(* IEC 61131-3 sources: plc-st-coding-agent/progress/evidence/f14_v10_full_20261113/jobs/custom_deepseek-v4pro (part 3) *)

(* ---- public-hard-05.raw_candidate_01.st ---- *)
FUNCTION_BLOCK MechanicalArmControl
VAR_INPUT
    ManualMode : BOOL;
    SingleStepMode : BOOL;
    SingleCycleMode : BOOL;
    ContinuousMode : BOOL;
    EmergencyStop : BOOL;
    Start : BOOL;
    DownButton : BOOL;
    UpButton : BOOL;
    LeftButton : BOOL;
    RightButton : BOOL;
    GripButton : BOOL;
    ReleaseButton : BOOL;
    DownLimitSwitch : BOOL;
    UpLimitSwitch : BOOL;
    LeftLimitSwitch : BOOL;
    RightLimitSwitch : BOOL;
    GripLimitSwitch : BOOL;
    ReleaseLimitSwitch : BOOL;
END_VAR
VAR_OUTPUT
    MoveDown : BOOL;
    MoveUp : BOOL;
    MoveLeft : BOOL;
    MoveRight : BOOL;
    ActivateGrip : BOOL;
    ActivateRelease : BOOL;
END_VAR
VAR
    local_StartRTrig : R_TRIG;
    local_StartEdge : BOOL;
    local_AutoActive : BOOL := FALSE;
    local_AutoStep : INT := 0;
    local_StepComplete : BOOL;
    local_DesiredMoveDown : BOOL;
    local_DesiredMoveUp : BOOL;
    local_DesiredMoveLeft : BOOL;
    local_DesiredMoveRight : BOOL;
    local_DesiredActivateGrip : BOOL;
    local_DesiredActivateRelease : BOOL;
END_VAR

(* ENGINEERING_CONTRACT
   Manual outputs: active in ManualMode while button=1 and limit=0;
   deactivate on button release, limit reached, or EmergencyStop=FALSE (PUB001, PUB005).
   SingleStep: Start edge begins current step; holds until limit; waits for next Start (PUB002, PUB003).
   SingleCycle: Start edge starts step0; automatic step advance on limit; stops after left (PUB003, PUB015-PUB017).
   Continuous: Start edge starts step0; automatically repeats after left (PUB004, PUB015-PUB017).
   E-stop: all outputs FALSE while EmergencyStop=FALSE; state frozen (PUB005).
   Auto steps 0..7: down,grip,up,right,down,release,up,left; completion via corresponding limit.
   Units/type: BOOL only; no timers; retained state local_AutoActive/local_AutoStep.
*)

(* CONTRACT_RULES [] *)

local_StartRTrig(CLK := Start);
local_StartEdge := local_StartRTrig.Q;

IF NOT EmergencyStop THEN
    MoveDown := FALSE;
    MoveUp := FALSE;
    MoveLeft := FALSE;
    MoveRight := FALSE;
    ActivateGrip := FALSE;
    ActivateRelease := FALSE;
    RETURN;
END_IF;

local_DesiredMoveDown := FALSE;
local_DesiredMoveUp := FALSE;
local_DesiredMoveLeft := FALSE;
local_DesiredMoveRight := FALSE;
local_DesiredActivateGrip := FALSE;
local_DesiredActivateRelease := FALSE;

IF ManualMode THEN
    IF DownButton AND NOT DownLimitSwitch THEN
        local_DesiredMoveDown := TRUE;
    END_IF;
    IF UpButton AND NOT UpLimitSwitch THEN
        local_DesiredMoveUp := TRUE;
    END_IF;
    IF LeftButton AND NOT LeftLimitSwitch THEN
        local_DesiredMoveLeft := TRUE;
    END_IF;
    IF RightButton AND NOT RightLimitSwitch THEN
        local_DesiredMoveRight := TRUE;
    END_IF;
    IF GripButton AND NOT GripLimitSwitch THEN
        local_DesiredActivateGrip := TRUE;
    END_IF;
    IF ReleaseButton AND NOT ReleaseLimitSwitch THEN
        local_DesiredActivateRelease := TRUE;
    END_IF;

ELSIF SingleStepMode OR SingleCycleMode OR ContinuousMode THEN
    IF SingleStepMode THEN
        IF local_StartEdge AND NOT local_AutoActive THEN
            local_AutoActive := TRUE;
        END_IF;

    ELSIF SingleCycleMode THEN
        IF local_StartEdge THEN
            local_AutoStep := 0;
            local_AutoActive := TRUE;
        END_IF;

    ELSIF ContinuousMode THEN
        IF local_StartEdge THEN
            local_AutoStep := 0;
            local_AutoActive := TRUE;
        END_IF;
    END_IF;

    IF local_AutoActive THEN
        CASE local_AutoStep OF
            0: local_DesiredMoveDown := NOT DownLimitSwitch;
            1: local_DesiredActivateGrip := NOT GripLimitSwitch;
            2: local_DesiredMoveUp := NOT UpLimitSwitch;
            3: local_DesiredMoveRight := NOT RightLimitSwitch;
            4: local_DesiredMoveDown := NOT DownLimitSwitch;
            5: local_DesiredActivateRelease := NOT ReleaseLimitSwitch;
            6: local_DesiredMoveUp := NOT UpLimitSwitch;
            7: local_DesiredMoveLeft := NOT LeftLimitSwitch;
        ELSE
            // no active output for invalid step
        END_CASE;
    END_IF;
END_IF;

MoveDown := local_DesiredMoveDown;
MoveUp := local_DesiredMoveUp;
MoveLeft := local_DesiredMoveLeft;
MoveRight := local_DesiredMoveRight;
ActivateGrip := local_DesiredActivateGrip;
ActivateRelease := local_DesiredActivateRelease;

IF SingleStepMode OR SingleCycleMode OR ContinuousMode THEN
    IF local_AutoActive THEN
        local_StepComplete := FALSE;

        IF (local_AutoStep = 0) OR (local_AutoStep = 4) THEN
            local_StepComplete := DownLimitSwitch;
        ELSIF (local_AutoStep = 1) THEN
            local_StepComplete := GripLimitSwitch;
        ELSIF (local_AutoStep = 2) OR (local_AutoStep = 6) THEN
            local_StepComplete := UpLimitSwitch;
        ELSIF (local_AutoStep = 3) THEN
            local_StepComplete := RightLimitSwitch;
        ELSIF (local_AutoStep = 5) THEN
            local_StepComplete := ReleaseLimitSwitch;
        ELSIF (local_AutoStep = 7) THEN
            local_StepComplete := LeftLimitSwitch;
        END_IF;

        IF local_StepComplete THEN
            IF SingleStepMode THEN
                local_AutoActive := FALSE;
                local_AutoStep := (local_AutoStep + 1) MOD 8;

            ELSIF SingleCycleMode THEN
                IF local_AutoStep < 7 THEN
                    local_AutoStep := local_AutoStep + 1;
                    // local_AutoActive remains TRUE
                ELSE
                    local_AutoActive := FALSE;
                    local_AutoStep := 0;
                END_IF;

            ELSIF ContinuousMode THEN
                local_AutoStep := (local_AutoStep + 1) MOD 8;
                local_AutoActive := TRUE;
            END_IF;
        END_IF;
    END_IF;
END_IF;

END_FUNCTION_BLOCK

(* ---- public-hard-05.raw_candidate_02.st ---- *)
FUNCTION_BLOCK MechanicalArmControl
VAR_INPUT
    ManualMode : BOOL;
    SingleStepMode : BOOL;
    SingleCycleMode : BOOL;
    ContinuousMode : BOOL;
    EmergencyStop : BOOL;
    Start : BOOL;
    DownButton : BOOL;
    UpButton : BOOL;
    LeftButton : BOOL;
    RightButton : BOOL;
    GripButton : BOOL;
    ReleaseButton : BOOL;
    DownLimitSwitch : BOOL;
    UpLimitSwitch : BOOL;
    LeftLimitSwitch : BOOL;
    RightLimitSwitch : BOOL;
    GripLimitSwitch : BOOL;
    ReleaseLimitSwitch : BOOL;
END_VAR
VAR_OUTPUT
    MoveDown : BOOL;
    MoveUp : BOOL;
    MoveLeft : BOOL;
    MoveRight : BOOL;
    ActivateGrip : BOOL;
    ActivateRelease : BOOL;
END_VAR
VAR
    local_StartRTrig : R_TRIG;
    local_StartEdge : BOOL;
    local_AutoActive : BOOL := FALSE;
    local_AutoStep : INT := 0;
    local_StepComplete : BOOL;
    local_DesiredMoveDown : BOOL;
    local_DesiredMoveUp : BOOL;
    local_DesiredMoveLeft : BOOL;
    local_DesiredMoveRight : BOOL;
    local_DesiredActivateGrip : BOOL;
    local_DesiredActivateRelease : BOOL;
END_VAR

(* ENGINEERING_CONTRACT
   Manual outputs: active in ManualMode while button=1 and limit=0;
   deactivate on button release, limit reached, or EmergencyStop=FALSE (PUB001, PUB005).
   SingleStep: Start edge begins current step; holds until limit; waits for next Start (PUB002, PUB003).
   SingleCycle: Start edge starts step0; automatic step advance on limit; stops after left (PUB003, PUB015-PUB017).
   Continuous: Start edge starts step0; automatically repeats after left (PUB004, PUB015-PUB017).
   E-stop: all outputs FALSE while EmergencyStop=FALSE; state frozen (PUB005).
   Auto steps 0..7: down,grip,up,right,down,release,up,left; completion via corresponding limit.
   Units/type: BOOL only; no timers; retained state local_AutoActive/local_AutoStep.
*)

(* CONTRACT_RULES [] *)

local_StartRTrig(CLK := Start);
local_StartEdge := local_StartRTrig.Q;

IF NOT EmergencyStop THEN
    MoveDown := FALSE;
    MoveUp := FALSE;
    MoveLeft := FALSE;
    MoveRight := FALSE;
    ActivateGrip := FALSE;
    ActivateRelease := FALSE;
    RETURN;
END_IF;

local_DesiredMoveDown := FALSE;
local_DesiredMoveUp := FALSE;
local_DesiredMoveLeft := FALSE;
local_DesiredMoveRight := FALSE;
local_DesiredActivateGrip := FALSE;
local_DesiredActivateRelease := FALSE;

IF ManualMode THEN
    IF DownButton AND NOT DownLimitSwitch THEN
        local_DesiredMoveDown := TRUE;
    END_IF;
    IF UpButton AND NOT UpLimitSwitch THEN
        local_DesiredMoveUp := TRUE;
    END_IF;
    IF LeftButton AND NOT LeftLimitSwitch THEN
        local_DesiredMoveLeft := TRUE;
    END_IF;
    IF RightButton AND NOT RightLimitSwitch THEN
        local_DesiredMoveRight := TRUE;
    END_IF;
    IF GripButton AND NOT GripLimitSwitch THEN
        local_DesiredActivateGrip := TRUE;
    END_IF;
    IF ReleaseButton AND NOT ReleaseLimitSwitch THEN
        local_DesiredActivateRelease := TRUE;
    END_IF;

ELSIF SingleStepMode OR SingleCycleMode OR ContinuousMode THEN
    IF SingleStepMode THEN
        IF local_StartEdge AND NOT local_AutoActive THEN
            local_AutoActive := TRUE;
        END_IF;

    ELSIF SingleCycleMode THEN
        IF local_StartEdge THEN
            local_AutoStep := 0;
            local_AutoActive := TRUE;
        END_IF;

    ELSIF ContinuousMode THEN
        IF local_StartEdge THEN
            local_AutoStep := 0;
            local_AutoActive := TRUE;
        END_IF;
    END_IF;

    IF local_AutoActive THEN
        CASE local_AutoStep OF
            0: local_DesiredMoveDown := NOT DownLimitSwitch;
            1: local_DesiredActivateGrip := NOT GripLimitSwitch;
            2: local_DesiredMoveUp := NOT UpLimitSwitch;
            3: local_DesiredMoveRight := NOT RightLimitSwitch;
            4: local_DesiredMoveDown := NOT DownLimitSwitch;
            5: local_DesiredActivateRelease := NOT ReleaseLimitSwitch;
            6: local_DesiredMoveUp := NOT UpLimitSwitch;
            7: local_DesiredMoveLeft := NOT LeftLimitSwitch;
        ELSE
            // no active output for invalid step
        END_CASE;
    END_IF;
END_IF;

MoveDown := local_DesiredMoveDown;
MoveUp := local_DesiredMoveUp;
MoveLeft := local_DesiredMoveLeft;
MoveRight := local_DesiredMoveRight;
ActivateGrip := local_DesiredActivateGrip;
ActivateRelease := local_DesiredActivateRelease;

IF SingleStepMode OR SingleCycleMode OR ContinuousMode THEN
    IF local_AutoActive THEN
        local_StepComplete := FALSE;

        IF (local_AutoStep = 0) OR (local_AutoStep = 4) THEN
            local_StepComplete := DownLimitSwitch;
        ELSIF (local_AutoStep = 1) THEN
            local_StepComplete := GripLimitSwitch;
        ELSIF (local_AutoStep = 2) OR (local_AutoStep = 6) THEN
            local_StepComplete := UpLimitSwitch;
        ELSIF (local_AutoStep = 3) THEN
            local_StepComplete := RightLimitSwitch;
        ELSIF (local_AutoStep = 5) THEN
            local_StepComplete := ReleaseLimitSwitch;
        ELSIF (local_AutoStep = 7) THEN
            local_StepComplete := LeftLimitSwitch;
        END_IF;

        IF local_StepComplete THEN
            IF SingleStepMode THEN
                local_AutoActive := FALSE;
                local_AutoStep := (local_AutoStep + 1) MOD 8;

            ELSIF SingleCycleMode THEN
                IF local_AutoStep < 7 THEN
                    local_AutoStep := local_AutoStep + 1;
                    (* local_AutoActive remains TRUE *)
                ELSE
                    local_AutoActive := FALSE;
                    local_AutoStep := 0;
                END_IF;

            ELSIF ContinuousMode THEN
                local_AutoStep := (local_AutoStep + 1) MOD 8;
                local_AutoActive := TRUE;
            END_IF;
        END_IF;
    END_IF;
END_IF;

END_FUNCTION_BLOCK

(* ---- public-hard-05.raw_candidate_03.st ---- *)
FUNCTION_BLOCK MechanicalArmControl
VAR_INPUT
    ManualMode : BOOL;
    SingleStepMode : BOOL;
    SingleCycleMode : BOOL;
    ContinuousMode : BOOL;
    EmergencyStop : BOOL;
    Start : BOOL;
    DownButton : BOOL;
    UpButton : BOOL;
    LeftButton : BOOL;
    RightButton : BOOL;
    GripButton : BOOL;
    ReleaseButton : BOOL;
    DownLimitSwitch : BOOL;
    UpLimitSwitch : BOOL;
    LeftLimitSwitch : BOOL;
    RightLimitSwitch : BOOL;
    GripLimitSwitch : BOOL;
    ReleaseLimitSwitch : BOOL;
END_VAR
VAR_OUTPUT
    MoveDown : BOOL;
    MoveUp : BOOL;
    MoveLeft : BOOL;
    MoveRight : BOOL;
    ActivateGrip : BOOL;
    ActivateRelease : BOOL;
END_VAR
VAR
    local_StartRTrig : R_TRIG;
    local_StartEdge : BOOL;
    local_AutoActive : BOOL := FALSE;
    local_AutoStep : INT := 0;
    local_StepComplete : BOOL;
    local_DesiredMoveDown : BOOL;
    local_DesiredMoveUp : BOOL;
    local_DesiredMoveLeft : BOOL;
    local_DesiredMoveRight : BOOL;
    local_DesiredActivateGrip : BOOL;
    local_DesiredActivateRelease : BOOL;
END_VAR

(* ENGINEERING_CONTRACT
   Manual outputs: active in ManualMode while button=1 and limit=0;
   deactivate on button release, limit reached, or EmergencyStop=FALSE (PUB001, PUB005).
   SingleStep: Start edge begins current step; holds until limit; waits for next Start (PUB002, PUB003).
   SingleCycle: Start edge starts step0; automatic step advance on limit; stops after left (PUB003, PUB015-PUB017).
   Continuous: Start edge starts step0; automatically repeats after left (PUB004, PUB015-PUB017).
   E-stop: all outputs FALSE while EmergencyStop=FALSE; state frozen (PUB005).
   Auto steps 0..7: down,grip,up,right,down,release,up,left; completion via corresponding limit.
   Units/type: BOOL only; no timers; retained state local_AutoActive/local_AutoStep.
*)

(* CONTRACT_RULES [] *)

local_StartRTrig(CLK := Start);
local_StartEdge := local_StartRTrig.Q;

(* Emergency stop has highest priority: immediately clear all outputs and return *)
IF NOT EmergencyStop THEN
    MoveDown := FALSE;
    MoveUp := FALSE;
    MoveLeft := FALSE;
    MoveRight := FALSE;
    ActivateGrip := FALSE;
    ActivateRelease := FALSE;
    RETURN;
END_IF;

(* Initialize desired outputs to FALSE *)
local_DesiredMoveDown := FALSE;
local_DesiredMoveUp := FALSE;
local_DesiredMoveLeft := FALSE;
local_DesiredMoveRight := FALSE;
local_DesiredActivateGrip := FALSE;
local_DesiredActivateRelease := FALSE;

IF ManualMode THEN
    (* Manual control: each action individually driven by its button and limit switch *)
    IF DownButton AND NOT DownLimitSwitch THEN
        local_DesiredMoveDown := TRUE;
    END_IF;
    IF UpButton AND NOT UpLimitSwitch THEN
        local_DesiredMoveUp := TRUE;
    END_IF;
    IF LeftButton AND NOT LeftLimitSwitch THEN
        local_DesiredMoveLeft := TRUE;
    END_IF;
    IF RightButton AND NOT RightLimitSwitch THEN
        local_DesiredMoveRight := TRUE;
    END_IF;
    IF GripButton AND NOT GripLimitSwitch THEN
        local_DesiredActivateGrip := TRUE;
    END_IF;
    IF ReleaseButton AND NOT ReleaseLimitSwitch THEN
        local_DesiredActivateRelease := TRUE;
    END_IF;

ELSIF SingleStepMode OR SingleCycleMode OR ContinuousMode THEN
    (* Automatic modes : single step, single cycle, continuous *)

    IF SingleStepMode THEN
        (* Activate on rising edge of Start only if not already active *)
        IF local_StartEdge AND NOT local_AutoActive THEN
            local_AutoActive := TRUE;
        END_IF;
    ELSIF SingleCycleMode THEN
        (* In single cycle, rising edge of Start resets sequence to step 0 and activates *)
        IF local_StartEdge THEN
            local_AutoStep := 0;
            local_AutoActive := TRUE;
        END_IF;
    ELSIF ContinuousMode THEN
        (* In continuous mode, rising edge of Start resets sequence to step 0 and activates *)
        IF local_StartEdge THEN
            local_AutoStep := 0;
            local_AutoActive := TRUE;
        END_IF;
    END_IF;

    IF local_AutoActive THEN
        CASE local_AutoStep OF
            0: local_DesiredMoveDown := NOT DownLimitSwitch;
            1: local_DesiredActivateGrip := NOT GripLimitSwitch;
            2: local_DesiredMoveUp := NOT UpLimitSwitch;
            3: local_DesiredMoveRight := NOT RightLimitSwitch;
            4: local_DesiredMoveDown := NOT DownLimitSwitch;
            5: local_DesiredActivateRelease := NOT ReleaseLimitSwitch;
            6: local_DesiredMoveUp := NOT UpLimitSwitch;
            7: local_DesiredMoveLeft := NOT LeftLimitSwitch;
        ELSE
            (* Invalid step: no desired movement *)
        END_CASE;
    END_IF;
END_IF;

(* Assign outputs from desired states *)
MoveDown := local_DesiredMoveDown;
MoveUp := local_DesiredMoveUp;
MoveLeft := local_DesiredMoveLeft;
MoveRight := local_DesiredMoveRight;
ActivateGrip := local_DesiredActivateGrip;
ActivateRelease := local_DesiredActivateRelease;

(* Handle step completion and transitions for automatic modes *)
IF SingleStepMode OR SingleCycleMode OR ContinuousMode THEN
    IF local_AutoActive THEN
        local_StepComplete := FALSE;

        IF local_AutoStep = 0 OR local_AutoStep = 4 THEN
            local_StepComplete := DownLimitSwitch;
        ELSIF local_AutoStep = 1 THEN
            local_StepComplete := GripLimitSwitch;
        ELSIF local_AutoStep = 2 OR local_AutoStep = 6 THEN
            local_StepComplete := UpLimitSwitch;
        ELSIF local_AutoStep = 3 THEN
            local_StepComplete := RightLimitSwitch;
        ELSIF local_AutoStep = 5 THEN
            local_StepComplete := ReleaseLimitSwitch;
        ELSIF local_AutoStep = 7 THEN
            local_StepComplete := LeftLimitSwitch;
        END_IF;

        IF local_StepComplete THEN
            IF SingleStepMode THEN
                (* Step finished: deactivate and advance step for next start *)
                local_AutoActive := FALSE;
                local_AutoStep := (local_AutoStep + 1) MOD 8;

            ELSIF SingleCycleMode THEN
                IF local_AutoStep < 7 THEN
                    (* Move to next step in sequence *)
                    local_AutoStep := local_AutoStep + 1;
                    (* local_AutoActive remains TRUE *)
                ELSE
                    (* Cycle complete: stop and reset for next start *)
                    local_AutoActive := FALSE;
                    local_AutoStep := 0;
                END_IF;

            ELSIF ContinuousMode THEN
                (* Automatically advance to next step and continue cycling *)
                local_AutoStep := (local_AutoStep + 1) MOD 8;
                local_AutoActive := TRUE;
            END_IF;
        END_IF;
    END_IF;
END_IF;

END_FUNCTION_BLOCK

(* ---- public-hard-05.raw_candidate_04.st ---- *)
FUNCTION_BLOCK MechanicalArmControl
VAR_INPUT
    ManualMode : BOOL;
    SingleStepMode : BOOL;
    SingleCycleMode : BOOL;
    ContinuousMode : BOOL;
    EmergencyStop : BOOL;
    Start : BOOL;
    DownButton : BOOL;
    UpButton : BOOL;
    LeftButton : BOOL;
    RightButton : BOOL;
    GripButton : BOOL;
    ReleaseButton : BOOL;
    DownLimitSwitch : BOOL;
    UpLimitSwitch : BOOL;
    LeftLimitSwitch : BOOL;
    RightLimitSwitch : BOOL;
    GripLimitSwitch : BOOL;
    ReleaseLimitSwitch : BOOL;
END_VAR
VAR_OUTPUT
    MoveDown : BOOL;
    MoveUp : BOOL;
    MoveLeft : BOOL;
    MoveRight : BOOL;
    ActivateGrip : BOOL;
    ActivateRelease : BOOL;
END_VAR
VAR
    local_StartRTrig : R_TRIG;
    local_StartEdge : BOOL;
    local_AutoActive : BOOL := FALSE;
    local_AutoStep : INT := 0;
    local_StepComplete : BOOL;
    local_DesiredMoveDown : BOOL;
    local_DesiredMoveUp : BOOL;
    local_DesiredMoveLeft : BOOL;
    local_DesiredMoveRight : BOOL;
    local_DesiredActivateGrip : BOOL;
    local_DesiredActivateRelease : BOOL;
END_VAR

(* ENGINEERING_CONTRACT
   Manual outputs: active in ManualMode while button=1 and limit=0;
   deactivate on button release, limit reached, or EmergencyStop=FALSE (PUB001, PUB005).
   SingleStep: Start edge begins current step; holds until limit; waits for next Start (PUB002, PUB003).
   SingleCycle: Start edge starts step0; automatic step advance on limit; stops after left (PUB003, PUB015-PUB017).
   Continuous: Start edge starts step0; automatically repeats after left (PUB004, PUB015-PUB017).
   E-stop: all outputs FALSE while EmergencyStop=FALSE; state frozen (PUB005).
   Auto steps 0..7: down,grip,up,right,down,release,up,left; completion via corresponding limit.
   Units/type: BOOL only; no timers; retained state local_AutoActive/local_AutoStep.
*)

(* CONTRACT_RULES [] *)

local_StartRTrig(CLK := Start);
local_StartEdge := local_StartRTrig.Q;

IF NOT EmergencyStop THEN
    MoveDown := FALSE;
    MoveUp := FALSE;
    MoveLeft := FALSE;
    MoveRight := FALSE;
    ActivateGrip := FALSE;
    ActivateRelease := FALSE;
    RETURN;
END_IF

local_DesiredMoveDown := FALSE;
local_DesiredMoveUp := FALSE;
local_DesiredMoveLeft := FALSE;
local_DesiredMoveRight := FALSE;
local_DesiredActivateGrip := FALSE;
local_DesiredActivateRelease := FALSE;

IF ManualMode THEN
    IF DownButton AND NOT DownLimitSwitch THEN
        local_DesiredMoveDown := TRUE;
    END_IF
    IF UpButton AND NOT UpLimitSwitch THEN
        local_DesiredMoveUp := TRUE;
    END_IF
    IF LeftButton AND NOT LeftLimitSwitch THEN
        local_DesiredMoveLeft := TRUE;
    END_IF
    IF RightButton AND NOT RightLimitSwitch THEN
        local_DesiredMoveRight := TRUE;
    END_IF
    IF GripButton AND NOT GripLimitSwitch THEN
        local_DesiredActivateGrip := TRUE;
    END_IF
    IF ReleaseButton AND NOT ReleaseLimitSwitch THEN
        local_DesiredActivateRelease := TRUE;
    END_IF

ELSIF SingleStepMode OR SingleCycleMode OR ContinuousMode THEN
    IF SingleStepMode THEN
        IF local_StartEdge AND NOT local_AutoActive THEN
            local_AutoActive := TRUE;
        END_IF

    ELSIF SingleCycleMode THEN
        IF local_StartEdge THEN
            local_AutoStep := 0;
            local_AutoActive := TRUE;
        END_IF

    ELSIF ContinuousMode THEN
        IF local_StartEdge THEN
            local_AutoStep := 0;
            local_AutoActive := TRUE;
        END_IF
    END_IF

    IF local_AutoActive THEN
        CASE local_AutoStep OF
            0: local_DesiredMoveDown := NOT DownLimitSwitch;
            1: local_DesiredActivateGrip := NOT GripLimitSwitch;
            2: local_DesiredMoveUp := NOT UpLimitSwitch;
            3: local_DesiredMoveRight := NOT RightLimitSwitch;
            4: local_DesiredMoveDown := NOT DownLimitSwitch;
            5: local_DesiredActivateRelease := NOT ReleaseLimitSwitch;
            6: local_DesiredMoveUp := NOT UpLimitSwitch;
            7: local_DesiredMoveLeft := NOT LeftLimitSwitch;
        ELSE
            // no active output for invalid step
        END_CASE
    END_IF
END_IF

MoveDown := local_DesiredMoveDown;
MoveUp := local_DesiredMoveUp;
MoveLeft := local_DesiredMoveLeft;
MoveRight := local_DesiredMoveRight;
ActivateGrip := local_DesiredActivateGrip;
ActivateRelease := local_DesiredActivateRelease;

IF SingleStepMode OR SingleCycleMode OR ContinuousMode THEN
    IF local_AutoActive THEN
        local_StepComplete := FALSE;

        IF (local_AutoStep = 0) OR (local_AutoStep = 4) THEN
            local_StepComplete := DownLimitSwitch;
        ELSIF (local_AutoStep = 1) THEN
            local_StepComplete := GripLimitSwitch;
        ELSIF (local_AutoStep = 2) OR (local_AutoStep = 6) THEN
            local_StepComplete := UpLimitSwitch;
        ELSIF (local_AutoStep = 3) THEN
            local_StepComplete := RightLimitSwitch;
        ELSIF (local_AutoStep = 5) THEN
            local_StepComplete := ReleaseLimitSwitch;
        ELSIF (local_AutoStep = 7) THEN
            local_StepComplete := LeftLimitSwitch;
        END_IF

        IF local_StepComplete THEN
            IF SingleStepMode THEN
                local_AutoActive := FALSE;
                local_AutoStep := (local_AutoStep + 1) MOD 8;

            ELSIF SingleCycleMode THEN
                IF local_AutoStep < 7 THEN
                    local_AutoStep := local_AutoStep + 1;
                    // local_AutoActive remains TRUE
                ELSE
                    local_AutoActive := FALSE;
                    local_AutoStep := 0;
                END_IF

            ELSIF ContinuousMode THEN
                local_AutoStep := (local_AutoStep + 1) MOD 8;
                local_AutoActive := TRUE;
            END_IF
        END_IF
    END_IF
END_IF

END_FUNCTION_BLOCK

(* ---- public-hard-06.candidate_01.st ---- *)
TYPE ProductionState : (IDLE, TO_WASH, AT_WASH, TO_WEIGHT, AT_WEIGHT, TO_FIRING, AT_FIRING, TO_OUTPUT, AT_OUTPUT, REJECTING) := IDLE;
END_TYPE;

(* ENGINEERING_CONTRACT
Manual forward/reverse: Mode=0; active when corresponding button true and other false; simultaneous => both false (PUB002).
Auto forward: active in TO_WASH/TO_WEIGHT/TO_FIRING/TO_OUTPUT; deasserted when target sensor activates; retained while moving (PUB003-PUB005).
Auto stop: AT_WASH/AT_WEIGHT/AT_FIRING/AT_OUTPUT wait for complete signal or removal; no edge detection (PUB003-PUB006).
kick: active when unqualified at weighing station after weightComplete; held until SensorWeight false; manual clears (PUB003).
CompletionLight: active while SensorOutput true in AT_OUTPUT; deasserted on SensorOutput false or manual (PUB006).
firingTemp: computed on qualified weight: 500+(weight-100)*0.5 for weight 100..200; retained through firing/output; cleared otherwise/manual (PUB003).
State: non-retain; starts IDLE; transitions by public sensors/signals; unspecified behavior if sensors overlap or mode changes mid-cycle.
*)
(* CONTRACT_RULES [] *)

FUNCTION_BLOCK ProductionControl
VAR_INPUT
    Mode : BOOL;
    ForwardButton : BOOL;
    ReverseButton : BOOL;
    SensorFeed : BOOL;
    SensorWash : BOOL;
    SensorWeight : BOOL;
    SensorFiring : BOOL;
    SensorOutput : BOOL;
    washComplete : BOOL;
    weightComplete : BOOL;
    weight : REAL;
    firingComplete : BOOL;
END_VAR
VAR_OUTPUT
    MotorForward : BOOL;
    MotorReverse : BOOL;
    kick : BOOL;
    CompletionLight : BOOL;
    firingTemp : REAL;
END_VAR
VAR
    state : ProductionState := ProductionState#IDLE;
    local_temp : REAL := 0.0;
END_VAR

IF Mode THEN
    (* Automatic mode *)
    MotorReverse := FALSE;
    CASE state OF
        ProductionState#IDLE:
            MotorForward := FALSE;
            kick := FALSE;
            firingTemp := 0.0;
            CompletionLight := FALSE;
            IF SensorFeed THEN
                state := ProductionState#TO_WASH;
            END_IF;

        ProductionState#TO_WASH:
            MotorForward := TRUE;
            kick := FALSE;
            firingTemp := 0.0;
            CompletionLight := FALSE;
            IF SensorWash THEN
                MotorForward := FALSE;
                state := ProductionState#AT_WASH;
            END_IF;

        ProductionState#AT_WASH:
            MotorForward := FALSE;
            kick := FALSE;
            firingTemp := 0.0;
            CompletionLight := FALSE;
            IF washComplete THEN
                MotorForward := TRUE;
                state := ProductionState#TO_WEIGHT;
            END_IF;

        ProductionState#TO_WEIGHT:
            MotorForward := TRUE;
            kick := FALSE;
            firingTemp := 0.0;
            CompletionLight := FALSE;
            IF SensorWeight THEN
                MotorForward := FALSE;
                state := ProductionState#AT_WEIGHT;
            END_IF;

        ProductionState#AT_WEIGHT:
            MotorForward := FALSE;
            kick := FALSE;
            firingTemp := 0.0;
            CompletionLight := FALSE;
            IF weightComplete THEN
                IF (weight >= 100.0) AND (weight <= 200.0) THEN
                    local_temp := 500.0 + (weight - 100.0) * 0.5;
                    firingTemp := local_temp;
                    state := ProductionState#TO_FIRING;
                ELSE
                    firingTemp := 0.0;
                    kick := TRUE;
                    state := ProductionState#REJECTING;
                END_IF;
            END_IF;

        ProductionState#REJECTING:
            MotorForward := FALSE;
            kick := TRUE;
            firingTemp := 0.0;
            CompletionLight := FALSE;
            IF NOT SensorWeight THEN
                kick := FALSE;
                state := ProductionState#IDLE;
            END_IF;

        ProductionState#TO_FIRING:
            MotorForward := TRUE;
            kick := FALSE;
            firingTemp := local_temp;
            CompletionLight := FALSE;
            IF SensorFiring THEN
                MotorForward := FALSE;
                state := ProductionState#AT_FIRING;
            END_IF;

        ProductionState#AT_FIRING:
            MotorForward := FALSE;
            kick := FALSE;
            firingTemp := local_temp;
            CompletionLight := FALSE;
            IF firingComplete THEN
                MotorForward := TRUE;
                state := ProductionState#TO_OUTPUT;
            END_IF;

        ProductionState#TO_OUTPUT:
            MotorForward := TRUE;
            kick := FALSE;
            firingTemp := local_temp;
            CompletionLight := FALSE;
            IF SensorOutput THEN
                MotorForward := FALSE;
                state := ProductionState#AT_OUTPUT;
            END_IF;

        ProductionState#AT_OUTPUT:
            MotorForward := FALSE;
            kick := FALSE;
            firingTemp := local_temp;
            CompletionLight := TRUE;
            IF NOT SensorOutput THEN
                CompletionLight := FALSE;
                state := ProductionState#IDLE;
            END_IF;
    END_CASE;
ELSE
    (* Manual mode *)
    MotorForward := FALSE;
    MotorReverse := FALSE;
    kick := FALSE;
    CompletionLight := FALSE;
    firingTemp := 0.0;

    IF ForwardButton AND NOT ReverseButton THEN
        MotorForward := TRUE;
        MotorReverse := FALSE;
    ELSIF ReverseButton AND NOT ForwardButton THEN
        MotorForward := FALSE;
        MotorReverse := TRUE;
    ELSE
        MotorForward := FALSE;
        MotorReverse := FALSE;
    END_IF;
END_IF;

END_FUNCTION_BLOCK

(* ---- public-hard-06.candidate_02.st ---- *)
TYPE ProductionState : (IDLE, TO_WASH, AT_WASH, TO_WEIGHT, AT_WEIGHT, TO_FIRING, AT_FIRING, TO_OUTPUT, AT_OUTPUT, REJECTING) := IDLE;
END_TYPE;

(* ENGINEERING_CONTRACT
Manual forward/reverse: Mode=0; active when corresponding button true and other false; simultaneous => both false (PUB002).
Auto forward: active in TO_WASH/TO_WEIGHT/TO_FIRING/TO_OUTPUT; deasserted when target sensor activates; retained while moving (PUB003-PUB005).
Auto stop: AT_WASH/AT_WEIGHT/AT_FIRING/AT_OUTPUT wait for complete signal or removal; no edge detection (PUB003-PUB006).
kick: active when unqualified at weighing station after weightComplete; held until SensorWeight false; manual clears (PUB003).
CompletionLight: active while SensorOutput true in AT_OUTPUT; deasserted on SensorOutput false or manual (PUB006).
firingTemp: computed on qualified weight: 500+(weight-100)*0.5 for weight 100..200; retained through firing/output; cleared otherwise/manual (PUB003).
State: non-retain; starts IDLE; transitions by public sensors/signals; unspecified behavior if sensors overlap or mode changes mid-cycle.
*)
(* CONTRACT_RULES [] *)

FUNCTION_BLOCK ProductionControl
VAR_INPUT
    Mode : BOOL;
    ForwardButton : BOOL;
    ReverseButton : BOOL;
    SensorFeed : BOOL;
    SensorWash : BOOL;
    SensorWeight : BOOL;
    SensorFiring : BOOL;
    SensorOutput : BOOL;
    washComplete : BOOL;
    weightComplete : BOOL;
    weight : REAL;
    firingComplete : BOOL;
END_VAR
VAR_OUTPUT
    MotorForward : BOOL;
    MotorReverse : BOOL;
    kick : BOOL;
    CompletionLight : BOOL;
    firingTemp : REAL;
END_VAR
VAR
    state : ProductionState := ProductionState.IDLE;
    local_temp : REAL := 0.0;
END_VAR

IF Mode THEN
    (* Automatic mode *)
    MotorReverse := FALSE;
    CASE state OF
        IDLE:
            MotorForward := FALSE;
            kick := FALSE;
            firingTemp := 0.0;
            CompletionLight := FALSE;
            IF SensorFeed THEN
                state := ProductionState.TO_WASH;
            END_IF;

        TO_WASH:
            MotorForward := TRUE;
            kick := FALSE;
            firingTemp := 0.0;
            CompletionLight := FALSE;
            IF SensorWash THEN
                MotorForward := FALSE;
                state := ProductionState.AT_WASH;
            END_IF;

        AT_WASH:
            MotorForward := FALSE;
            kick := FALSE;
            firingTemp := 0.0;
            CompletionLight := FALSE;
            IF washComplete THEN
                MotorForward := TRUE;
                state := ProductionState.TO_WEIGHT;
            END_IF;

        TO_WEIGHT:
            MotorForward := TRUE;
            kick := FALSE;
            firingTemp := 0.0;
            CompletionLight := FALSE;
            IF SensorWeight THEN
                MotorForward := FALSE;
                state := ProductionState.AT_WEIGHT;
            END_IF;

        AT_WEIGHT:
            MotorForward := FALSE;
            kick := FALSE;
            firingTemp := 0.0;
            CompletionLight := FALSE;
            IF weightComplete THEN
                IF (weight >= 100.0) AND (weight <= 200.0) THEN
                    local_temp := 500.0 + (weight - 100.0) * 0.5;
                    firingTemp := local_temp;
                    MotorForward := TRUE; (* immediate forward on qualification *)
                    state := ProductionState.TO_FIRING;
                ELSE
                    firingTemp := 0.0;
                    kick := TRUE;
                    state := ProductionState.REJECTING;
                END_IF;
            END_IF;

        REJECTING:
            MotorForward := FALSE;
            kick := TRUE;
            firingTemp := 0.0;
            CompletionLight := FALSE;
            IF NOT SensorWeight THEN
                kick := FALSE;
                state := ProductionState.IDLE;
            END_IF;

        TO_FIRING:
            MotorForward := TRUE;
            kick := FALSE;
            firingTemp := local_temp;
            CompletionLight := FALSE;
            IF SensorFiring THEN
                MotorForward := FALSE;
                state := ProductionState.AT_FIRING;
            END_IF;

        AT_FIRING:
            MotorForward := FALSE;
            kick := FALSE;
            firingTemp := local_temp;
            CompletionLight := FALSE;
            IF firingComplete THEN
                MotorForward := TRUE;
                state := ProductionState.TO_OUTPUT;
            END_IF;

        TO_OUTPUT:
            MotorForward := TRUE;
            kick := FALSE;
            firingTemp := local_temp;
            CompletionLight := FALSE;
            IF SensorOutput THEN
                MotorForward := FALSE;
                state := ProductionState.AT_OUTPUT;
            END_IF;

        AT_OUTPUT:
            MotorForward := FALSE;
            kick := FALSE;
            firingTemp := local_temp;
            CompletionLight := TRUE;
            IF NOT SensorOutput THEN
                CompletionLight := FALSE;
                state := ProductionState.IDLE;
            END_IF;
    END_CASE;
ELSE
    (* Manual mode *)
    MotorForward := FALSE;
    MotorReverse := FALSE;
    kick := FALSE;
    CompletionLight := FALSE;
    firingTemp := 0.0;

    IF ForwardButton AND NOT ReverseButton THEN
        MotorForward := TRUE;
        MotorReverse := FALSE;
    ELSIF ReverseButton AND NOT ForwardButton THEN
        MotorForward := FALSE;
        MotorReverse := TRUE;
    ELSE
        MotorForward := FALSE;
        MotorReverse := FALSE;
    END_IF;
END_IF;

END_FUNCTION_BLOCK

(* ---- public-hard-06.candidate_03.st ---- *)
TYPE ProductionState : (IDLE, TO_WASH, AT_WASH, TO_WEIGHT, AT_WEIGHT, TO_FIRING, AT_FIRING, TO_OUTPUT, AT_OUTPUT, REJECTING) := IDLE;
END_TYPE;

(* ENGINEERING_CONTRACT
Manual forward/reverse: Mode=0; active when corresponding button true and other false; simultaneous => both false (PUB002).
Auto forward: active in TO_WASH/TO_WEIGHT/TO_FIRING/TO_OUTPUT; deasserted when target sensor activates; retained while moving (PUB003-PUB005).
Auto stop: AT_WASH/AT_WEIGHT/AT_FIRING/AT_OUTPUT wait for complete signal or removal; no edge detection (PUB003-PUB006).
kick: active when unqualified at weighing station after weightComplete; held until SensorWeight false; manual clears (PUB003).
CompletionLight: active while SensorOutput true in AT_OUTPUT; deasserted on SensorOutput false or manual (PUB006).
firingTemp: computed on qualified weight: 500+(weight-100)*0.5 for weight 100..200; retained through firing/output; cleared otherwise/manual (PUB003).
State: non-retain; starts IDLE; transitions by public sensors/signals; unspecified behavior if sensors overlap or mode changes mid-cycle.
Same-scan: outputs are recomputed after every state transition in the same invocation.
*)
(* CONTRACT_RULES [] *)

FUNCTION_BLOCK ProductionControl
VAR_INPUT
    Mode : BOOL;
    ForwardButton : BOOL;
    ReverseButton : BOOL;
    SensorFeed : BOOL;
    SensorWash : BOOL;
    SensorWeight : BOOL;
    SensorFiring : BOOL;
    SensorOutput : BOOL;
    washComplete : BOOL;
    weightComplete : BOOL;
    weight : REAL;
    firingComplete : BOOL;
END_VAR
VAR_OUTPUT
    MotorForward : BOOL;
    MotorReverse : BOOL;
    kick : BOOL;
    CompletionLight : BOOL;
    firingTemp : REAL;
END_VAR
VAR
    state : ProductionState := ProductionState.IDLE;
    local_temp : REAL := 0.0;
END_VAR

IF Mode THEN
    (* Automatic mode *)
    MotorReverse := FALSE;

    (* State transition logic *)
    CASE state OF
        IDLE:
            IF SensorFeed THEN
                state := ProductionState.TO_WASH;
            END_IF;

        TO_WASH:
            IF SensorWash THEN
                state := ProductionState.AT_WASH;
            END_IF;

        AT_WASH:
            IF washComplete THEN
                state := ProductionState.TO_WEIGHT;
            END_IF;

        TO_WEIGHT:
            IF SensorWeight THEN
                state := ProductionState.AT_WEIGHT;
            END_IF;

        AT_WEIGHT:
            IF weightComplete THEN
                IF (weight >= 100.0) AND (weight <= 200.0) THEN
                    local_temp := 500.0 + (weight - 100.0) * 0.5;
                    state := ProductionState.TO_FIRING;
                ELSE
                    state := ProductionState.REJECTING;
                END_IF;
            END_IF;

        REJECTING:
            IF NOT SensorWeight THEN
                state := ProductionState.IDLE;
            END_IF;

        TO_FIRING:
            IF SensorFiring THEN
                state := ProductionState.AT_FIRING;
            END_IF;

        AT_FIRING:
            IF firingComplete THEN
                state := ProductionState.TO_OUTPUT;
            END_IF;

        TO_OUTPUT:
            IF SensorOutput THEN
                state := ProductionState.AT_OUTPUT;
            END_IF;

        AT_OUTPUT:
            IF NOT SensorOutput THEN
                state := ProductionState.IDLE;
            END_IF;
    END_CASE;

    (* Compute outputs from current state after transitions *)
    MotorForward := FALSE;
    kick := FALSE;
    CompletionLight := FALSE;
    firingTemp := 0.0;

    CASE state OF
        TO_WASH, TO_WEIGHT, TO_FIRING, TO_OUTPUT:
            MotorForward := TRUE;
    END_CASE;

    IF (state = AT_OUTPUT) AND SensorOutput THEN
        CompletionLight := TRUE;
    END_IF;

    IF (state = REJECTING) AND SensorWeight THEN
        kick := TRUE;
    END_IF;

    IF (state = TO_FIRING) OR (state = AT_FIRING) OR (state = TO_OUTPUT) OR (state = AT_OUTPUT) THEN
        firingTemp := local_temp;
    END_IF;

ELSE
    (* Manual mode *)
    MotorForward := FALSE;
    MotorReverse := FALSE;
    kick := FALSE;
    CompletionLight := FALSE;
    firingTemp := 0.0;

    IF ForwardButton AND NOT ReverseButton THEN
        MotorForward := TRUE;
    ELSIF ReverseButton AND NOT ForwardButton THEN
        MotorReverse := TRUE;
    ELSE
        MotorForward := FALSE;
        MotorReverse := FALSE;
    END_IF;
END_IF;

END_FUNCTION_BLOCK

(* ---- public-hard-06.candidate_04.st ---- *)
TYPE ProductionState : (IDLE, TO_WASH, AT_WASH, TO_WEIGHT, AT_WEIGHT, TO_FIRING, AT_FIRING, TO_OUTPUT, AT_OUTPUT, REJECTING) := IDLE;
END_TYPE;

(* ENGINEERING_CONTRACT
Manual forward/reverse: Mode=0; active when corresponding button true and other false; simultaneous => both false (PUB002).
Auto forward: active in TO_WASH/TO_WEIGHT/TO_FIRING/TO_OUTPUT; deasserted when target sensor activates; retained while moving (PUB003-PUB005).
Auto stop: AT_WASH/AT_WEIGHT/AT_FIRING/AT_OUTPUT wait for complete signal or removal; no edge detection (PUB003-PUB006).
kick: active when unqualified at weighing station after weightComplete; held until SensorWeight false; manual clears (PUB003).
CompletionLight: active while SensorOutput true in AT_OUTPUT; deasserted on SensorOutput false or manual (PUB006).
firingTemp: computed on qualified weight: 500+(weight-100)*0.5 for weight 100..200; retained through firing/output and after product removal until next qualification or manual (PUB003).
State: non-retain; starts IDLE; transitions by public sensors/signals; unspecified behavior if sensors overlap or mode changes mid-cycle.
Same-scan: outputs are recomputed after every state transition in the same invocation.
*)
(* CONTRACT_RULES [] *)

FUNCTION_BLOCK ProductionControl
VAR_INPUT
    Mode : BOOL;
    ForwardButton : BOOL;
    ReverseButton : BOOL;
    SensorFeed : BOOL;
    SensorWash : BOOL;
    SensorWeight : BOOL;
    SensorFiring : BOOL;
    SensorOutput : BOOL;
    washComplete : BOOL;
    weightComplete : BOOL;
    weight : REAL;
    firingComplete : BOOL;
END_VAR
VAR_OUTPUT
    MotorForward : BOOL;
    MotorReverse : BOOL;
    kick : BOOL;
    CompletionLight : BOOL;
    firingTemp : REAL;
END_VAR
VAR
    state : ProductionState := ProductionState.IDLE;
    local_temp : REAL := 0.0;
END_VAR

IF Mode THEN
    (* Automatic mode *)
    MotorReverse := FALSE;

    (* State transition logic *)
    CASE state OF
        IDLE:
            IF SensorFeed THEN
                state := ProductionState.TO_WASH;
            END_IF;

        TO_WASH:
            IF SensorWash THEN
                state := ProductionState.AT_WASH;
            END_IF;

        AT_WASH:
            IF washComplete THEN
                state := ProductionState.TO_WEIGHT;
            END_IF;

        TO_WEIGHT:
            IF SensorWeight THEN
                state := ProductionState.AT_WEIGHT;
            END_IF;

        AT_WEIGHT:
            IF weightComplete THEN
                IF (weight >= 100.0) AND (weight <= 200.0) THEN
                    local_temp := 500.0 + (weight - 100.0) * 0.5;
                    state := ProductionState.TO_FIRING;
                ELSE
                    firingTemp := 0.0; (* clear previous temperature on unqualified *)
                    state := ProductionState.REJECTING;
                END_IF;
            END_IF;

        REJECTING:
            IF NOT SensorWeight THEN
                state := ProductionState.IDLE;
            END_IF;

        TO_FIRING:
            IF SensorFiring THEN
                state := ProductionState.AT_FIRING;
            END_IF;

        AT_FIRING:
            IF firingComplete THEN
                state := ProductionState.TO_OUTPUT;
            END_IF;

        TO_OUTPUT:
            IF SensorOutput THEN
                state := ProductionState.AT_OUTPUT;
            END_IF;

        AT_OUTPUT:
            IF NOT SensorOutput THEN
                state := ProductionState.IDLE;
            END_IF;
    END_CASE;

    (* Compute outputs after transitions *)
    MotorForward := FALSE;
    kick := FALSE;
    CompletionLight := FALSE;
    (* firingTemp intentionally not globally reset; retains last qualified value unless cleared by manual/unqualified *)

    CASE state OF
        TO_WASH, TO_WEIGHT, TO_FIRING, TO_OUTPUT:
            MotorForward := TRUE;
    END_CASE;

    IF (state = AT_OUTPUT) AND SensorOutput THEN
        CompletionLight := TRUE;
    END_IF;

    IF (state = REJECTING) THEN
        kick := TRUE;
    END_IF;

    IF (state = TO_FIRING) OR (state = AT_FIRING) OR (state = TO_OUTPUT) OR (state = AT_OUTPUT) THEN
        firingTemp := local_temp;
    END_IF;

ELSE
    (* Manual mode *)
    MotorForward := FALSE;
    MotorReverse := FALSE;
    kick := FALSE;
    CompletionLight := FALSE;
    firingTemp := 0.0;

    IF ForwardButton AND NOT ReverseButton THEN
        MotorForward := TRUE;
    ELSIF ReverseButton AND NOT ForwardButton THEN
        MotorReverse := TRUE;
    ELSE
        MotorForward := FALSE;
        MotorReverse := FALSE;
    END_IF;
END_IF;

END_FUNCTION_BLOCK

(* ---- public-hard-06.raw_candidate_01.st ---- *)
TYPE ProductionState : (IDLE, TO_WASH, AT_WASH, TO_WEIGHT, AT_WEIGHT, TO_FIRING, AT_FIRING, TO_OUTPUT, AT_OUTPUT, REJECTING) := IDLE;
END_TYPE

(* ENGINEERING_CONTRACT
Manual forward/reverse: Mode=0; active when corresponding button true and other false; simultaneous => both false (PUB002).
Auto forward: active in TO_WASH/TO_WEIGHT/TO_FIRING/TO_OUTPUT; deasserted when target sensor activates; retained while moving (PUB003-PUB005).
Auto stop: AT_WASH/AT_WEIGHT/AT_FIRING/AT_OUTPUT wait for complete signal or removal; no edge detection (PUB003-PUB006).
kick: active when unqualified at weighing station after weightComplete; held until SensorWeight false; manual clears (PUB003).
CompletionLight: active while SensorOutput true in AT_OUTPUT; deasserted on SensorOutput false or manual (PUB006).
firingTemp: computed on qualified weight: 500+(weight-100)*0.5 for weight 100..200; retained through firing/output; cleared otherwise/manual (PUB003).
State: non-retain; starts IDLE; transitions by public sensors/signals; unspecified behavior if sensors overlap or mode changes mid-cycle.
*)
(* CONTRACT_RULES [] *)

FUNCTION_BLOCK ProductionControl
VAR_INPUT
    Mode : BOOL;
    ForwardButton : BOOL;
    ReverseButton : BOOL;
    SensorFeed : BOOL;
    SensorWash : BOOL;
    SensorWeight : BOOL;
    SensorFiring : BOOL;
    SensorOutput : BOOL;
    washComplete : BOOL;
    weightComplete : BOOL;
    weight : REAL;
    firingComplete : BOOL;
END_VAR
VAR_OUTPUT
    MotorForward : BOOL;
    MotorReverse : BOOL;
    kick : BOOL;
    CompletionLight : BOOL;
    firingTemp : REAL;
END_VAR
VAR
    state : ProductionState := ProductionState#IDLE;
    local_temp : REAL := 0.0;
END_VAR

IF Mode THEN
    (* Automatic mode *)
    MotorReverse := FALSE;
    CASE state OF
        ProductionState#IDLE:
            MotorForward := FALSE;
            kick := FALSE;
            firingTemp := 0.0;
            CompletionLight := FALSE;
            IF SensorFeed THEN
                state := ProductionState#TO_WASH;
            END_IF;

        ProductionState#TO_WASH:
            MotorForward := TRUE;
            kick := FALSE;
            firingTemp := 0.0;
            CompletionLight := FALSE;
            IF SensorWash THEN
                MotorForward := FALSE;
                state := ProductionState#AT_WASH;
            END_IF;

        ProductionState#AT_WASH:
            MotorForward := FALSE;
            kick := FALSE;
            firingTemp := 0.0;
            CompletionLight := FALSE;
            IF washComplete THEN
                MotorForward := TRUE;
                state := ProductionState#TO_WEIGHT;
            END_IF;

        ProductionState#TO_WEIGHT:
            MotorForward := TRUE;
            kick := FALSE;
            firingTemp := 0.0;
            CompletionLight := FALSE;
            IF SensorWeight THEN
                MotorForward := FALSE;
                state := ProductionState#AT_WEIGHT;
            END_IF;

        ProductionState#AT_WEIGHT:
            MotorForward := FALSE;
            kick := FALSE;
            firingTemp := 0.0;
            CompletionLight := FALSE;
            IF weightComplete THEN
                IF (weight >= 100.0) AND (weight <= 200.0) THEN
                    local_temp := 500.0 + (weight - 100.0) * 0.5;
                    firingTemp := local_temp;
                    state := ProductionState#TO_FIRING;
                ELSE
                    firingTemp := 0.0;
                    kick := TRUE;
                    state := ProductionState#REJECTING;
                END_IF;
            END_IF;

        ProductionState#REJECTING:
            MotorForward := FALSE;
            kick := TRUE;
            firingTemp := 0.0;
            CompletionLight := FALSE;
            IF NOT SensorWeight THEN
                kick := FALSE;
                state := ProductionState#IDLE;
            END_IF;

        ProductionState#TO_FIRING:
            MotorForward := TRUE;
            kick := FALSE;
            firingTemp := local_temp;
            CompletionLight := FALSE;
            IF SensorFiring THEN
                MotorForward := FALSE;
                state := ProductionState#AT_FIRING;
            END_IF;

        ProductionState#AT_FIRING:
            MotorForward := FALSE;
            kick := FALSE;
            firingTemp := local_temp;
            CompletionLight := FALSE;
            IF firingComplete THEN
                MotorForward := TRUE;
                state := ProductionState#TO_OUTPUT;
            END_IF;

        ProductionState#TO_OUTPUT:
            MotorForward := TRUE;
            kick := FALSE;
            firingTemp := local_temp;
            CompletionLight := FALSE;
            IF SensorOutput THEN
                MotorForward := FALSE;
                state := ProductionState#AT_OUTPUT;
            END_IF;

        ProductionState#AT_OUTPUT:
            MotorForward := FALSE;
            kick := FALSE;
            firingTemp := local_temp;
            CompletionLight := TRUE;
            IF NOT SensorOutput THEN
                CompletionLight := FALSE;
                state := ProductionState#IDLE;
            END_IF;
    END_CASE;
ELSE
    (* Manual mode *)
    MotorForward := FALSE;
    MotorReverse := FALSE;
    kick := FALSE;
    CompletionLight := FALSE;
    firingTemp := 0.0;

    IF ForwardButton AND NOT ReverseButton THEN
        MotorForward := TRUE;
        MotorReverse := FALSE;
    ELSIF ReverseButton AND NOT ForwardButton THEN
        MotorForward := FALSE;
        MotorReverse := TRUE;
    ELSE
        MotorForward := FALSE;
        MotorReverse := FALSE;
    END_IF;
END_IF;

END_FUNCTION_BLOCK

(* ---- public-hard-06.raw_candidate_02.st ---- *)
TYPE ProductionState : (IDLE, TO_WASH, AT_WASH, TO_WEIGHT, AT_WEIGHT, TO_FIRING, AT_FIRING, TO_OUTPUT, AT_OUTPUT, REJECTING) := IDLE;
END_TYPE;

(* ENGINEERING_CONTRACT
Manual forward/reverse: Mode=0; active when corresponding button true and other false; simultaneous => both false (PUB002).
Auto forward: active in TO_WASH/TO_WEIGHT/TO_FIRING/TO_OUTPUT; deasserted when target sensor activates; retained while moving (PUB003-PUB005).
Auto stop: AT_WASH/AT_WEIGHT/AT_FIRING/AT_OUTPUT wait for complete signal or removal; no edge detection (PUB003-PUB006).
kick: active when unqualified at weighing station after weightComplete; held until SensorWeight false; manual clears (PUB003).
CompletionLight: active while SensorOutput true in AT_OUTPUT; deasserted on SensorOutput false or manual (PUB006).
firingTemp: computed on qualified weight: 500+(weight-100)*0.5 for weight 100..200; retained through firing/output; cleared otherwise/manual (PUB003).
State: non-retain; starts IDLE; transitions by public sensors/signals; unspecified behavior if sensors overlap or mode changes mid-cycle.
*)
(* CONTRACT_RULES [] *)

FUNCTION_BLOCK ProductionControl
VAR_INPUT
    Mode : BOOL;
    ForwardButton : BOOL;
    ReverseButton : BOOL;
    SensorFeed : BOOL;
    SensorWash : BOOL;
    SensorWeight : BOOL;
    SensorFiring : BOOL;
    SensorOutput : BOOL;
    washComplete : BOOL;
    weightComplete : BOOL;
    weight : REAL;
    firingComplete : BOOL;
END_VAR
VAR_OUTPUT
    MotorForward : BOOL;
    MotorReverse : BOOL;
    kick : BOOL;
    CompletionLight : BOOL;
    firingTemp : REAL;
END_VAR
VAR
    state : ProductionState := ProductionState.IDLE;
    local_temp : REAL := 0.0;
END_VAR

IF Mode THEN
    (* Automatic mode *)
    MotorReverse := FALSE;
    CASE state OF
        IDLE:
            MotorForward := FALSE;
            kick := FALSE;
            firingTemp := 0.0;
            CompletionLight := FALSE;
            IF SensorFeed THEN
                state := ProductionState.TO_WASH;
            END_IF;

        TO_WASH:
            MotorForward := TRUE;
            kick := FALSE;
            firingTemp := 0.0;
            CompletionLight := FALSE;
            IF SensorWash THEN
                MotorForward := FALSE;
                state := ProductionState.AT_WASH;
            END_IF;

        AT_WASH:
            MotorForward := FALSE;
            kick := FALSE;
            firingTemp := 0.0;
            CompletionLight := FALSE;
            IF washComplete THEN
                MotorForward := TRUE;
                state := ProductionState.TO_WEIGHT;
            END_IF;

        TO_WEIGHT:
            MotorForward := TRUE;
            kick := FALSE;
            firingTemp := 0.0;
            CompletionLight := FALSE;
            IF SensorWeight THEN
                MotorForward := FALSE;
                state := ProductionState.AT_WEIGHT;
            END_IF;

        AT_WEIGHT:
            MotorForward := FALSE;
            kick := FALSE;
            firingTemp := 0.0;
            CompletionLight := FALSE;
            IF weightComplete THEN
                IF (weight >= 100.0) AND (weight <= 200.0) THEN
                    local_temp := 500.0 + (weight - 100.0) * 0.5;
                    firingTemp := local_temp;
                    MotorForward := TRUE; (* immediate forward on qualification *)
                    state := ProductionState.TO_FIRING;
                ELSE
                    firingTemp := 0.0;
                    kick := TRUE;
                    state := ProductionState.REJECTING;
                END_IF;
            END_IF;

        REJECTING:
            MotorForward := FALSE;
            kick := TRUE;
            firingTemp := 0.0;
            CompletionLight := FALSE;
            IF NOT SensorWeight THEN
                kick := FALSE;
                state := ProductionState.IDLE;
            END_IF;

        TO_FIRING:
            MotorForward := TRUE;
            kick := FALSE;
            firingTemp := local_temp;
            CompletionLight := FALSE;
            IF SensorFiring THEN
                MotorForward := FALSE;
                state := ProductionState.AT_FIRING;
            END_IF;

        AT_FIRING:
            MotorForward := FALSE;
            kick := FALSE;
            firingTemp := local_temp;
            CompletionLight := FALSE;
            IF firingComplete THEN
                MotorForward := TRUE;
                state := ProductionState.TO_OUTPUT;
            END_IF;

        TO_OUTPUT:
            MotorForward := TRUE;
            kick := FALSE;
            firingTemp := local_temp;
            CompletionLight := FALSE;
            IF SensorOutput THEN
                MotorForward := FALSE;
                state := ProductionState.AT_OUTPUT;
            END_IF;

        AT_OUTPUT:
            MotorForward := FALSE;
            kick := FALSE;
            firingTemp := local_temp;
            CompletionLight := TRUE;
            IF NOT SensorOutput THEN
                CompletionLight := FALSE;
                state := ProductionState.IDLE;
            END_IF;
    END_CASE;
ELSE
    (* Manual mode *)
    MotorForward := FALSE;
    MotorReverse := FALSE;
    kick := FALSE;
    CompletionLight := FALSE;
    firingTemp := 0.0;

    IF ForwardButton AND NOT ReverseButton THEN
        MotorForward := TRUE;
        MotorReverse := FALSE;
    ELSIF ReverseButton AND NOT ForwardButton THEN
        MotorForward := FALSE;
        MotorReverse := TRUE;
    ELSE
        MotorForward := FALSE;
        MotorReverse := FALSE;
    END_IF;
END_IF;

END_FUNCTION_BLOCK

(* ---- public-hard-06.raw_candidate_03.st ---- *)
TYPE ProductionState : (IDLE, TO_WASH, AT_WASH, TO_WEIGHT, AT_WEIGHT, TO_FIRING, AT_FIRING, TO_OUTPUT, AT_OUTPUT, REJECTING) := IDLE;
END_TYPE;

(* ENGINEERING_CONTRACT
Manual forward/reverse: Mode=0; active when corresponding button true and other false; simultaneous => both false (PUB002).
Auto forward: active in TO_WASH/TO_WEIGHT/TO_FIRING/TO_OUTPUT; deasserted when target sensor activates; retained while moving (PUB003-PUB005).
Auto stop: AT_WASH/AT_WEIGHT/AT_FIRING/AT_OUTPUT wait for complete signal or removal; no edge detection (PUB003-PUB006).
kick: active when unqualified at weighing station after weightComplete; held until SensorWeight false; manual clears (PUB003).
CompletionLight: active while SensorOutput true in AT_OUTPUT; deasserted on SensorOutput false or manual (PUB006).
firingTemp: computed on qualified weight: 500+(weight-100)*0.5 for weight 100..200; retained through firing/output; cleared otherwise/manual (PUB003).
State: non-retain; starts IDLE; transitions by public sensors/signals; unspecified behavior if sensors overlap or mode changes mid-cycle.
Same-scan: outputs are recomputed after every state transition in the same invocation.
*)
(* CONTRACT_RULES [] *)

FUNCTION_BLOCK ProductionControl
VAR_INPUT
    Mode : BOOL;
    ForwardButton : BOOL;
    ReverseButton : BOOL;
    SensorFeed : BOOL;
    SensorWash : BOOL;
    SensorWeight : BOOL;
    SensorFiring : BOOL;
    SensorOutput : BOOL;
    washComplete : BOOL;
    weightComplete : BOOL;
    weight : REAL;
    firingComplete : BOOL;
END_VAR
VAR_OUTPUT
    MotorForward : BOOL;
    MotorReverse : BOOL;
    kick : BOOL;
    CompletionLight : BOOL;
    firingTemp : REAL;
END_VAR
VAR
    state : ProductionState := ProductionState.IDLE;
    local_temp : REAL := 0.0;
END_VAR

IF Mode THEN
    (* Automatic mode *)
    MotorReverse := FALSE;

    (* State transition logic *)
    CASE state OF
        IDLE:
            IF SensorFeed THEN
                state := ProductionState.TO_WASH;
            END_IF;

        TO_WASH:
            IF SensorWash THEN
                state := ProductionState.AT_WASH;
            END_IF;

        AT_WASH:
            IF washComplete THEN
                state := ProductionState.TO_WEIGHT;
            END_IF;

        TO_WEIGHT:
            IF SensorWeight THEN
                state := ProductionState.AT_WEIGHT;
            END_IF;

        AT_WEIGHT:
            IF weightComplete THEN
                IF (weight >= 100.0) AND (weight <= 200.0) THEN
                    local_temp := 500.0 + (weight - 100.0) * 0.5;
                    state := ProductionState.TO_FIRING;
                ELSE
                    state := ProductionState.REJECTING;
                END_IF;
            END_IF;

        REJECTING:
            IF NOT SensorWeight THEN
                state := ProductionState.IDLE;
            END_IF;

        TO_FIRING:
            IF SensorFiring THEN
                state := ProductionState.AT_FIRING;
            END_IF;

        AT_FIRING:
            IF firingComplete THEN
                state := ProductionState.TO_OUTPUT;
            END_IF;

        TO_OUTPUT:
            IF SensorOutput THEN
                state := ProductionState.AT_OUTPUT;
            END_IF;

        AT_OUTPUT:
            IF NOT SensorOutput THEN
                state := ProductionState.IDLE;
            END_IF;
    END_CASE;

    (* Compute outputs from current state after transitions *)
    MotorForward := FALSE;
    kick := FALSE;
    CompletionLight := FALSE;
    firingTemp := 0.0;

    CASE state OF
        TO_WASH, TO_WEIGHT, TO_FIRING, TO_OUTPUT:
            MotorForward := TRUE;
    END_CASE;

    IF (state = AT_OUTPUT) AND SensorOutput THEN
        CompletionLight := TRUE;
    END_IF;

    IF (state = REJECTING) AND SensorWeight THEN
        kick := TRUE;
    END_IF;

    IF (state = TO_FIRING) OR (state = AT_FIRING) OR (state = TO_OUTPUT) OR (state = AT_OUTPUT) THEN
        firingTemp := local_temp;
    END_IF;

ELSE
    (* Manual mode *)
    MotorForward := FALSE;
    MotorReverse := FALSE;
    kick := FALSE;
    CompletionLight := FALSE;
    firingTemp := 0.0;

    IF ForwardButton AND NOT ReverseButton THEN
        MotorForward := TRUE;
    ELSIF ReverseButton AND NOT ForwardButton THEN
        MotorReverse := TRUE;
    ELSE
        MotorForward := FALSE;
        MotorReverse := FALSE;
    END_IF;
END_IF;

END_FUNCTION_BLOCK

(* ---- public-hard-06.raw_candidate_04.st ---- *)
TYPE ProductionState : (IDLE, TO_WASH, AT_WASH, TO_WEIGHT, AT_WEIGHT, TO_FIRING, AT_FIRING, TO_OUTPUT, AT_OUTPUT, REJECTING) := IDLE;
END_TYPE;

(* ENGINEERING_CONTRACT
Manual forward/reverse: Mode=0; active when corresponding button true and other false; simultaneous => both false (PUB002).
Auto forward: active in TO_WASH/TO_WEIGHT/TO_FIRING/TO_OUTPUT; deasserted when target sensor activates; retained while moving (PUB003-PUB005).
Auto stop: AT_WASH/AT_WEIGHT/AT_FIRING/AT_OUTPUT wait for complete signal or removal; no edge detection (PUB003-PUB006).
kick: active when unqualified at weighing station after weightComplete; held until SensorWeight false; manual clears (PUB003).
CompletionLight: active while SensorOutput true in AT_OUTPUT; deasserted on SensorOutput false or manual (PUB006).
firingTemp: computed on qualified weight: 500+(weight-100)*0.5 for weight 100..200; retained through firing/output and after product removal until next qualification or manual (PUB003).
State: non-retain; starts IDLE; transitions by public sensors/signals; unspecified behavior if sensors overlap or mode changes mid-cycle.
Same-scan: outputs are recomputed after every state transition in the same invocation.
*)
(* CONTRACT_RULES [] *)

FUNCTION_BLOCK ProductionControl
VAR_INPUT
    Mode : BOOL;
    ForwardButton : BOOL;
    ReverseButton : BOOL;
    SensorFeed : BOOL;
    SensorWash : BOOL;
    SensorWeight : BOOL;
    SensorFiring : BOOL;
    SensorOutput : BOOL;
    washComplete : BOOL;
    weightComplete : BOOL;
    weight : REAL;
    firingComplete : BOOL;
END_VAR
VAR_OUTPUT
    MotorForward : BOOL;
    MotorReverse : BOOL;
    kick : BOOL;
    CompletionLight : BOOL;
    firingTemp : REAL;
END_VAR
VAR
    state : ProductionState := ProductionState.IDLE;
    local_temp : REAL := 0.0;
END_VAR

IF Mode THEN
    (* Automatic mode *)
    MotorReverse := FALSE;

    (* State transition logic *)
    CASE state OF
        IDLE:
            IF SensorFeed THEN
                state := ProductionState.TO_WASH;
            END_IF;

        TO_WASH:
            IF SensorWash THEN
                state := ProductionState.AT_WASH;
            END_IF;

        AT_WASH:
            IF washComplete THEN
                state := ProductionState.TO_WEIGHT;
            END_IF;

        TO_WEIGHT:
            IF SensorWeight THEN
                state := ProductionState.AT_WEIGHT;
            END_IF;

        AT_WEIGHT:
            IF weightComplete THEN
                IF (weight >= 100.0) AND (weight <= 200.0) THEN
                    local_temp := 500.0 + (weight - 100.0) * 0.5;
                    state := ProductionState.TO_FIRING;
                ELSE
                    firingTemp := 0.0; (* clear previous temperature on unqualified *)
                    state := ProductionState.REJECTING;
                END_IF;
            END_IF;

        REJECTING:
            IF NOT SensorWeight THEN
                state := ProductionState.IDLE;
            END_IF;

        TO_FIRING:
            IF SensorFiring THEN
                state := ProductionState.AT_FIRING;
            END_IF;

        AT_FIRING:
            IF firingComplete THEN
                state := ProductionState.TO_OUTPUT;
            END_IF;

        TO_OUTPUT:
            IF SensorOutput THEN
                state := ProductionState.AT_OUTPUT;
            END_IF;

        AT_OUTPUT:
            IF NOT SensorOutput THEN
                state := ProductionState.IDLE;
            END_IF;
    END_CASE;

    (* Compute outputs after transitions *)
    MotorForward := FALSE;
    kick := FALSE;
    CompletionLight := FALSE;
    (* firingTemp intentionally not globally reset; retains last qualified value unless cleared by manual/unqualified *)

    CASE state OF
        TO_WASH, TO_WEIGHT, TO_FIRING, TO_OUTPUT:
            MotorForward := TRUE;
    END_CASE;

    IF (state = AT_OUTPUT) AND SensorOutput THEN
        CompletionLight := TRUE;
    END_IF;

    IF (state = REJECTING) THEN
        kick := TRUE;
    END_IF;

    IF (state = TO_FIRING) OR (state = AT_FIRING) OR (state = TO_OUTPUT) OR (state = AT_OUTPUT) THEN
        firingTemp := local_temp;
    END_IF;

ELSE
    (* Manual mode *)
    MotorForward := FALSE;
    MotorReverse := FALSE;
    kick := FALSE;
    CompletionLight := FALSE;
    firingTemp := 0.0;

    IF ForwardButton AND NOT ReverseButton THEN
        MotorForward := TRUE;
    ELSIF ReverseButton AND NOT ForwardButton THEN
        MotorReverse := TRUE;
    ELSE
        MotorForward := FALSE;
        MotorReverse := FALSE;
    END_IF;
END_IF;

END_FUNCTION_BLOCK

(* ---- public-medium-01.candidate_01.st ---- *)
TYPE ST_Pump :
STRUCT
    priority : INT;
    selection : BOOL;
    RunComd : BOOL;
END_STRUCT
END_TYPE;

FUNCTION_BLOCK MultiPumpSwitchingControl
VAR_INPUT
    mode : BOOL;
    start : BOOL;
    stop : BOOL;
END_VAR
VAR_IN_OUT
    pumpGroup : ARRAY[1..5] OF ST_Pump;
END_VAR
VAR
    tmp_runEnable : BOOL;
    tmp_i : INT;
    tmp_j : INT;
    tmp_higher : INT;
    tmp_equal_before : INT;
    tmp_selected : ARRAY[1..5] OF BOOL;
END_VAR

(* ENGINEERING_CONTRACT
   Mode/selection: mode=FALSE => manual set = pumpGroup[i].selection; mode=TRUE => auto set = top-3 priority values, tie lower index (PUB001, PUB003).
   Run command activation: start=TRUE with stop=FALSE latches tmp_runEnable=TRUE (PUB002).
   Retention/latch: tmp_runEnable holds after start until stop; each pump RunComd follows current mode/selection and tmp_runEnable every scan (PUB002).
   Stop/reset: stop=TRUE clears tmp_runEnable and all RunComd, same-scan priority over start and mode computation (PUB004).
   Boundaries: priority INT, exactly 3 pumps selected in auto, tie lower array index unspecified interpretation; only RunComd is written.
*)

(* CONTRACT_RULES [] *)

IF stop THEN
    tmp_runEnable := FALSE;
    FOR tmp_i := 1 TO 5 DO
        pumpGroup[tmp_i].RunComd := FALSE;
    END_FOR;
    RETURN;
END_IF;

IF start THEN
    tmp_runEnable := TRUE;
END_IF;

IF mode THEN
    FOR tmp_i := 1 TO 5 DO
        tmp_higher := 0;
        tmp_equal_before := 0;
        FOR tmp_j := 1 TO 5 DO
            IF pumpGroup[tmp_j].priority > pumpGroup[tmp_i].priority THEN
                tmp_higher := tmp_higher + 1;
            ELSIF (tmp_j < tmp_i) AND (pumpGroup[tmp_j].priority = pumpGroup[tmp_i].priority) THEN
                tmp_equal_before := tmp_equal_before + 1;
            END_IF;
        END_FOR;
        tmp_selected[tmp_i] := ((tmp_higher + tmp_equal_before) < 3);
    END_FOR;
    FOR tmp_i := 1 TO 5 DO
        pumpGroup[tmp_i].RunComd := tmp_runEnable AND tmp_selected[tmp_i];
    END_FOR;
ELSE
    FOR tmp_i := 1 TO 5 DO
        pumpGroup[tmp_i].RunComd := tmp_runEnable AND pumpGroup[tmp_i].selection;
    END_FOR;
END_IF;

END_FUNCTION_BLOCK

(* ---- public-medium-01.candidate_02.st ---- *)
TYPE ST_Pump :
STRUCT
    priority : INT;
    selection : BOOL;
    RunComd : BOOL;
END_STRUCT
END_TYPE;

FUNCTION_BLOCK MultiPumpSwitchingControl
VAR_INPUT
    mode : BOOL;
    start : BOOL;
    stop : BOOL;
END_VAR
VAR_IN_OUT
    pumpGroup : ARRAY[1..5] OF ST_Pump;
END_VAR
VAR
    tmp_runEnable : BOOL;
    tmp_i : INT;
    tmp_j : INT;
    tmp_higher : INT;
    tmp_equal_before : INT;
    tmp_selected : ARRAY[1..5] OF BOOL;
    tmp_startR : R_TRIG;
END_VAR

(* ENGINEERING_CONTRACT
   Mode/selection: mode=FALSE => manual set = pumpGroup[i].selection;
                   mode=TRUE  => auto set = top-3 priority values, tie lower index (PUB001, PUB003).
   Run command activation: rising edge of start when stop=FALSE latches tmp_runEnable=TRUE.
                           Start held after stop does not restart until a new rising edge.
   Retention/latch: tmp_runEnable holds after start until stop; each pump RunComd follows
                    current mode/selection and tmp_runEnable every scan (PUB002).
   Stop/reset: stop=TRUE clears tmp_runEnable and all RunComd, same-scan priority
               over start and mode computation (PUB004).
   Boundaries: priority INT, exactly 3 pumps selected in auto, tie lower index
               unspecified interpretation; only RunComd is written.
*)

(* CONTRACT_RULES [] *)

tmp_startR(CLK := start);

IF stop THEN
    tmp_runEnable := FALSE;
    FOR tmp_i := 1 TO 5 DO
        pumpGroup[tmp_i].RunComd := FALSE;
    END_FOR;
    RETURN;
END_IF;

IF tmp_startR.Q THEN
    tmp_runEnable := TRUE;
END_IF;

IF mode THEN
    FOR tmp_i := 1 TO 5 DO
        tmp_higher := 0;
        tmp_equal_before := 0;
        FOR tmp_j := 1 TO 5 DO
            IF pumpGroup[tmp_j].priority > pumpGroup[tmp_i].priority THEN
                tmp_higher := tmp_higher + 1;
            ELSIF (tmp_j < tmp_i) AND (pumpGroup[tmp_j].priority = pumpGroup[tmp_i].priority) THEN
                tmp_equal_before := tmp_equal_before + 1;
            END_IF;
        END_FOR;
        tmp_selected[tmp_i] := ((tmp_higher + tmp_equal_before) < 3);
    END_FOR;
    FOR tmp_i := 1 TO 5 DO
        pumpGroup[tmp_i].RunComd := tmp_runEnable AND tmp_selected[tmp_i];
    END_FOR;
ELSE
    FOR tmp_i := 1 TO 5 DO
        pumpGroup[tmp_i].RunComd := tmp_runEnable AND pumpGroup[tmp_i].selection;
    END_FOR;
END_IF;

END_FUNCTION_BLOCK

(* ---- public-medium-01.candidate_03.st ---- *)
TYPE ST_Pump :
STRUCT
    priority : INT;      (* Larger value = higher priority. Read-only to FB. *)
    selection : BOOL;    (* Manual-selection state. Read-only to FB. *)
    RunComd : BOOL;      (* Written by FB. TRUE = run, FALSE = stop. *)
END_STRUCT
END_TYPE;

FUNCTION_BLOCK MultiPumpSwitchingControl
VAR_INPUT
    mode  : BOOL;  (* FALSE = Manual, TRUE = Automatic *)
    start : BOOL;  (* Start button - rising-edge triggered *)
    stop  : BOOL;  (* Stop button - level sensitive, overrides start *)
END_VAR
VAR_IN_OUT
    pumpGroup : ARRAY[1..5] OF ST_Pump; (* Read priority/selection, write RunComd only *)
END_VAR
VAR
    tmp_runEnable      : BOOL;                    (* Latched run command state *)
    tmp_start_ris      : R_TRIG;                  (* Rising-edge detector for start *)
    tmp_i              : INT;
    tmp_j              : INT;
    tmp_higher         : INT;                     (* Number of pumps with strictly higher priority *)
    tmp_equal_before   : INT;                     (* Equal priority pumps with lower array index *)
    tmp_selected       : ARRAY[1..5] OF BOOL;     (* Automatic top-3 selection set *)
END_VAR

(* ENGINEERING_CONTRACT
   mode: FALSE=manual set = pumpGroup[i].selection; TRUE=auto set = top-3 priority values,
         ties resolved toward lower array index. Larger priority = higher priority.
   start: rising-edge latch, holds tmp_runEnable TRUE until stop.
   stop: level-sensitive, immediate priority over start and mode; clears latch and all RunComd.
   outputs: RunComd = tmp_runEnable AND selected/auto-selected for each pump.
   same-scan: stop wins over start; mode change immediately recomputes active set.
   boundaries: priority INT, exactly 3 pumps selected in auto, tie lower index.
*)

(* CONTRACT_RULES [] *)

(* Update start-edge memory every scan, even when stop is active,
   so a held start cannot false-trigger after stop is released. *)
tmp_start_ris(CLK := start);

IF stop THEN
    tmp_runEnable := FALSE;
    FOR tmp_i := 1 TO 5 DO
        pumpGroup[tmp_i].RunComd := FALSE;
    END_FOR;
    RETURN;
END_IF;

IF tmp_start_ris.Q THEN
    tmp_runEnable := TRUE;
END_IF;

IF mode THEN
    (* Automatic mode: select exactly 3 pumps with highest priority,
       lower array index used for ties. *)
    FOR tmp_i := 1 TO 5 DO
        tmp_higher := 0;
        tmp_equal_before := 0;
        FOR tmp_j := 1 TO 5 DO
            IF pumpGroup[tmp_j].priority > pumpGroup[tmp_i].priority THEN
                tmp_higher := tmp_higher + 1;
            ELSIF (tmp_j < tmp_i) AND (pumpGroup[tmp_j].priority = pumpGroup[tmp_i].priority) THEN
                tmp_equal_before := tmp_equal_before + 1;
            END_IF;
        END_FOR;
        tmp_selected[tmp_i] := ((tmp_higher + tmp_equal_before) < 3);
    END_FOR;

    FOR tmp_i := 1 TO 5 DO
        pumpGroup[tmp_i].RunComd := tmp_runEnable AND tmp_selected[tmp_i];
    END_FOR;
ELSE
    (* Manual mode: use each pump's manual selection. *)
    FOR tmp_i := 1 TO 5 DO
        pumpGroup[tmp_i].RunComd := tmp_runEnable AND pumpGroup[tmp_i].selection;
    END_FOR;
END_IF;

END_FUNCTION_BLOCK

(* ---- public-medium-01.candidate_04.st ---- *)
TYPE ST_Pump :
STRUCT
    priority : INT;
    selection : BOOL;
    RunComd : BOOL;
END_STRUCT
END_TYPE;

FUNCTION_BLOCK MultiPumpSwitchingControl
VAR_INPUT
    mode : BOOL;
    start : BOOL;
    stop : BOOL;
END_VAR
VAR_IN_OUT
    pumpGroup : ARRAY[1..5] OF ST_Pump;
END_VAR
VAR
    tmp_runEnable : BOOL;
    tmp_i : INT;
    tmp_j : INT;
    tmp_higher : INT;
    tmp_equal_before : INT;
    tmp_selected : ARRAY[1..5] OF BOOL;
    tmp_startRTrig : R_TRIG;
END_VAR

(* ENGINEERING_CONTRACT
   State tmp_runEnable: activation = rising edge of start while stop=FALSE; hold until stop; reset by stop.
   A start edge occurring while stop=TRUE is consumed and must be re-pressed after stop clears.
   RunComd group: activation = tmp_runEnable AND (manual selection OR auto top-3).
   stop has same-scan priority: clears tmp_runEnable and all RunComd before any start/mode logic.
   Auto selection: exactly 3 pumps; larger priority wins; equal priority tie by lower array index (unspecified).
   Manual selection: pumpGroup[i].selection directly gates RunComd while tmp_runEnable.
   Only RunComd is written; priority and selection are read-only.
*)

(* CONTRACT_RULES [] *)

tmp_startRTrig(CLK := start);

IF stop THEN
    tmp_runEnable := FALSE;
    FOR tmp_i := 1 TO 5 DO
        pumpGroup[tmp_i].RunComd := FALSE;
    END_FOR;
    RETURN;
END_IF;

IF tmp_startRTrig.Q THEN
    tmp_runEnable := TRUE;
END_IF;

IF mode THEN
    FOR tmp_i := 1 TO 5 DO
        tmp_higher := 0;
        tmp_equal_before := 0;
        FOR tmp_j := 1 TO 5 DO
            IF pumpGroup[tmp_j].priority > pumpGroup[tmp_i].priority THEN
                tmp_higher := tmp_higher + 1;
            ELSIF (tmp_j < tmp_i) AND (pumpGroup[tmp_j].priority = pumpGroup[tmp_i].priority) THEN
                tmp_equal_before := tmp_equal_before + 1;
            END_IF;
        END_FOR;
        tmp_selected[tmp_i] := ((tmp_higher + tmp_equal_before) < 3);
    END_FOR;

    FOR tmp_i := 1 TO 5 DO
        pumpGroup[tmp_i].RunComd := tmp_runEnable AND tmp_selected[tmp_i];
    END_FOR;
ELSE
    FOR tmp_i := 1 TO 5 DO
        pumpGroup[tmp_i].RunComd := tmp_runEnable AND pumpGroup[tmp_i].selection;
    END_FOR;
END_IF;

END_FUNCTION_BLOCK

(* ---- public-medium-01.raw_candidate_01.st ---- *)
TYPE ST_Pump :
STRUCT
    priority : INT;
    selection : BOOL;
    RunComd : BOOL;
END_STRUCT
END_TYPE

FUNCTION_BLOCK MultiPumpSwitchingControl
VAR_INPUT
    mode : BOOL;
    start : BOOL;
    stop : BOOL;
END_VAR
VAR_IN_OUT
    pumpGroup : ARRAY[1..5] OF ST_Pump;
END_VAR
VAR
    tmp_runEnable : BOOL;
    tmp_i : INT;
    tmp_j : INT;
    tmp_higher : INT;
    tmp_equal_before : INT;
    tmp_selected : ARRAY[1..5] OF BOOL;
END_VAR

(* ENGINEERING_CONTRACT
   Mode/selection: mode=FALSE => manual set = pumpGroup[i].selection; mode=TRUE => auto set = top-3 priority values, tie lower index (PUB001, PUB003).
   Run command activation: start=TRUE with stop=FALSE latches tmp_runEnable=TRUE (PUB002).
   Retention/latch: tmp_runEnable holds after start until stop; each pump RunComd follows current mode/selection and tmp_runEnable every scan (PUB002).
   Stop/reset: stop=TRUE clears tmp_runEnable and all RunComd, same-scan priority over start and mode computation (PUB004).
   Boundaries: priority INT, exactly 3 pumps selected in auto, tie lower array index unspecified interpretation; only RunComd is written.
*)

(* CONTRACT_RULES [] *)

IF stop THEN
    tmp_runEnable := FALSE;
    FOR tmp_i := 1 TO 5 DO
        pumpGroup[tmp_i].RunComd := FALSE;
    END_FOR;
    RETURN;
END_IF;

IF start THEN
    tmp_runEnable := TRUE;
END_IF;

IF mode THEN
    FOR tmp_i := 1 TO 5 DO
        tmp_higher := 0;
        tmp_equal_before := 0;
        FOR tmp_j := 1 TO 5 DO
            IF pumpGroup[tmp_j].priority > pumpGroup[tmp_i].priority THEN
                tmp_higher := tmp_higher + 1;
            ELSIF (tmp_j < tmp_i) AND (pumpGroup[tmp_j].priority = pumpGroup[tmp_i].priority) THEN
                tmp_equal_before := tmp_equal_before + 1;
            END_IF;
        END_FOR;
        tmp_selected[tmp_i] := ((tmp_higher + tmp_equal_before) < 3);
    END_FOR;
    FOR tmp_i := 1 TO 5 DO
        pumpGroup[tmp_i].RunComd := tmp_runEnable AND tmp_selected[tmp_i];
    END_FOR;
ELSE
    FOR tmp_i := 1 TO 5 DO
        pumpGroup[tmp_i].RunComd := tmp_runEnable AND pumpGroup[tmp_i].selection;
    END_FOR;
END_IF;

END_FUNCTION_BLOCK

(* ---- public-medium-01.raw_candidate_02.st ---- *)
TYPE ST_Pump :
STRUCT
    priority : INT;
    selection : BOOL;
    RunComd : BOOL;
END_STRUCT
END_TYPE;

FUNCTION_BLOCK MultiPumpSwitchingControl
VAR_INPUT
    mode : BOOL;
    start : BOOL;
    stop : BOOL;
END_VAR
VAR_IN_OUT
    pumpGroup : ARRAY[1..5] OF ST_Pump;
END_VAR
VAR
    tmp_runEnable : BOOL;
    tmp_i : INT;
    tmp_j : INT;
    tmp_higher : INT;
    tmp_equal_before : INT;
    tmp_selected : ARRAY[1..5] OF BOOL;
    tmp_startR : R_TRIG;
END_VAR

(* ENGINEERING_CONTRACT
   Mode/selection: mode=FALSE => manual set = pumpGroup[i].selection;
                   mode=TRUE  => auto set = top-3 priority values, tie lower index (PUB001, PUB003).
   Run command activation: rising edge of start when stop=FALSE latches tmp_runEnable=TRUE.
                           Start held after stop does not restart until a new rising edge.
   Retention/latch: tmp_runEnable holds after start until stop; each pump RunComd follows
                    current mode/selection and tmp_runEnable every scan (PUB002).
   Stop/reset: stop=TRUE clears tmp_runEnable and all RunComd, same-scan priority
               over start and mode computation (PUB004).
   Boundaries: priority INT, exactly 3 pumps selected in auto, tie lower index
               unspecified interpretation; only RunComd is written.
*)

(* CONTRACT_RULES [] *)

tmp_startR(CLK := start);

IF stop THEN
    tmp_runEnable := FALSE;
    FOR tmp_i := 1 TO 5 DO
        pumpGroup[tmp_i].RunComd := FALSE;
    END_FOR;
    RETURN;
END_IF;

IF tmp_startR.Q THEN
    tmp_runEnable := TRUE;
END_IF;

IF mode THEN
    FOR tmp_i := 1 TO 5 DO
        tmp_higher := 0;
        tmp_equal_before := 0;
        FOR tmp_j := 1 TO 5 DO
            IF pumpGroup[tmp_j].priority > pumpGroup[tmp_i].priority THEN
                tmp_higher := tmp_higher + 1;
            ELSIF (tmp_j < tmp_i) AND (pumpGroup[tmp_j].priority = pumpGroup[tmp_i].priority) THEN
                tmp_equal_before := tmp_equal_before + 1;
            END_IF;
        END_FOR;
        tmp_selected[tmp_i] := ((tmp_higher + tmp_equal_before) < 3);
    END_FOR;
    FOR tmp_i := 1 TO 5 DO
        pumpGroup[tmp_i].RunComd := tmp_runEnable AND tmp_selected[tmp_i];
    END_FOR;
ELSE
    FOR tmp_i := 1 TO 5 DO
        pumpGroup[tmp_i].RunComd := tmp_runEnable AND pumpGroup[tmp_i].selection;
    END_FOR;
END_IF;

END_FUNCTION_BLOCK

(* ---- public-medium-01.raw_candidate_03.st ---- *)
TYPE ST_Pump :
STRUCT
    priority : INT;      (* Larger value = higher priority. Read-only to FB. *)
    selection : BOOL;    (* Manual-selection state. Read-only to FB. *)
    RunComd : BOOL;      (* Written by FB. TRUE = run, FALSE = stop. *)
END_STRUCT
END_TYPE

FUNCTION_BLOCK MultiPumpSwitchingControl
VAR_INPUT
    mode  : BOOL;  (* FALSE = Manual, TRUE = Automatic *)
    start : BOOL;  (* Start button - rising-edge triggered *)
    stop  : BOOL;  (* Stop button - level sensitive, overrides start *)
END_VAR
VAR_IN_OUT
    pumpGroup : ARRAY[1..5] OF ST_Pump; (* Read priority/selection, write RunComd only *)
END_VAR
VAR
    tmp_runEnable      : BOOL;                    (* Latched run command state *)
    tmp_start_ris      : R_TRIG;                  (* Rising-edge detector for start *)
    tmp_i              : INT;
    tmp_j              : INT;
    tmp_higher         : INT;                     (* Number of pumps with strictly higher priority *)
    tmp_equal_before   : INT;                     (* Equal priority pumps with lower array index *)
    tmp_selected       : ARRAY[1..5] OF BOOL;     (* Automatic top-3 selection set *)
END_VAR

(* ENGINEERING_CONTRACT
   mode: FALSE=manual set = pumpGroup[i].selection; TRUE=auto set = top-3 priority values,
         ties resolved toward lower array index. Larger priority = higher priority.
   start: rising-edge latch, holds tmp_runEnable TRUE until stop.
   stop: level-sensitive, immediate priority over start and mode; clears latch and all RunComd.
   outputs: RunComd = tmp_runEnable AND selected/auto-selected for each pump.
   same-scan: stop wins over start; mode change immediately recomputes active set.
   boundaries: priority INT, exactly 3 pumps selected in auto, tie lower index.
*)

(* CONTRACT_RULES [] *)

(* Update start-edge memory every scan, even when stop is active,
   so a held start cannot false-trigger after stop is released. *)
tmp_start_ris(CLK := start);

IF stop THEN
    tmp_runEnable := FALSE;
    FOR tmp_i := 1 TO 5 DO
        pumpGroup[tmp_i].RunComd := FALSE;
    END_FOR;
    RETURN;
END_IF;

IF tmp_start_ris.Q THEN
    tmp_runEnable := TRUE;
END_IF;

IF mode THEN
    (* Automatic mode: select exactly 3 pumps with highest priority,
       lower array index used for ties. *)
    FOR tmp_i := 1 TO 5 DO
        tmp_higher := 0;
        tmp_equal_before := 0;
        FOR tmp_j := 1 TO 5 DO
            IF pumpGroup[tmp_j].priority > pumpGroup[tmp_i].priority THEN
                tmp_higher := tmp_higher + 1;
            ELSIF (tmp_j < tmp_i) AND (pumpGroup[tmp_j].priority = pumpGroup[tmp_i].priority) THEN
                tmp_equal_before := tmp_equal_before + 1;
            END_IF;
        END_FOR;
        tmp_selected[tmp_i] := ((tmp_higher + tmp_equal_before) < 3);
    END_FOR;

    FOR tmp_i := 1 TO 5 DO
        pumpGroup[tmp_i].RunComd := tmp_runEnable AND tmp_selected[tmp_i];
    END_FOR;
ELSE
    (* Manual mode: use each pump's manual selection. *)
    FOR tmp_i := 1 TO 5 DO
        pumpGroup[tmp_i].RunComd := tmp_runEnable AND pumpGroup[tmp_i].selection;
    END_FOR;
END_IF;

END_FUNCTION_BLOCK

(* ---- public-medium-01.raw_candidate_04.st ---- *)
TYPE ST_Pump :
STRUCT
    priority : INT;
    selection : BOOL;
    RunComd : BOOL;
END_STRUCT
END_TYPE

FUNCTION_BLOCK MultiPumpSwitchingControl
VAR_INPUT
    mode : BOOL;
    start : BOOL;
    stop : BOOL;
END_VAR
VAR_IN_OUT
    pumpGroup : ARRAY[1..5] OF ST_Pump;
END_VAR
VAR
    tmp_runEnable : BOOL;
    tmp_i : INT;
    tmp_j : INT;
    tmp_higher : INT;
    tmp_equal_before : INT;
    tmp_selected : ARRAY[1..5] OF BOOL;
    tmp_startRTrig : R_TRIG;
END_VAR

(* ENGINEERING_CONTRACT
   State tmp_runEnable: activation = rising edge of start while stop=FALSE; hold until stop; reset by stop.
   A start edge occurring while stop=TRUE is consumed and must be re-pressed after stop clears.
   RunComd group: activation = tmp_runEnable AND (manual selection OR auto top-3).
   stop has same-scan priority: clears tmp_runEnable and all RunComd before any start/mode logic.
   Auto selection: exactly 3 pumps; larger priority wins; equal priority tie by lower array index (unspecified).
   Manual selection: pumpGroup[i].selection directly gates RunComd while tmp_runEnable.
   Only RunComd is written; priority and selection are read-only.
*)

(* CONTRACT_RULES [] *)

tmp_startRTrig(CLK := start);

IF stop THEN
    tmp_runEnable := FALSE;
    FOR tmp_i := 1 TO 5 DO
        pumpGroup[tmp_i].RunComd := FALSE;
    END_FOR;
    RETURN;
END_IF;

IF tmp_startRTrig.Q THEN
    tmp_runEnable := TRUE;
END_IF;

IF mode THEN
    FOR tmp_i := 1 TO 5 DO
        tmp_higher := 0;
        tmp_equal_before := 0;
        FOR tmp_j := 1 TO 5 DO
            IF pumpGroup[tmp_j].priority > pumpGroup[tmp_i].priority THEN
                tmp_higher := tmp_higher + 1;
            ELSIF (tmp_j < tmp_i) AND (pumpGroup[tmp_j].priority = pumpGroup[tmp_i].priority) THEN
                tmp_equal_before := tmp_equal_before + 1;
            END_IF;
        END_FOR;
        tmp_selected[tmp_i] := ((tmp_higher + tmp_equal_before) < 3);
    END_FOR;

    FOR tmp_i := 1 TO 5 DO
        pumpGroup[tmp_i].RunComd := tmp_runEnable AND tmp_selected[tmp_i];
    END_FOR;
ELSE
    FOR tmp_i := 1 TO 5 DO
        pumpGroup[tmp_i].RunComd := tmp_runEnable AND pumpGroup[tmp_i].selection;
    END_FOR;
END_IF;

END_FUNCTION_BLOCK

(* ---- public-medium-02.candidate_01.st ---- *)
TYPE ST_AnalogChannel :
STRUCT
    enable : BOOL;
    hiLIM : REAL;
    loLIM : REAL;
    bipolar : BOOL;
    measuringMode : INT;
    retVal : WORD;
    outputValue : REAL;
END_STRUCT
END_TYPE;

(*
ENGINEERING_CONTRACT
Activation: process first count ordinal channels, count >= 0, clamped to min array lengths.
Enable: only channels[].enable = TRUE is evaluated; disabled rows retain previous retVal/outputValue.
retVal: for enabled rows write WORD#0 on success; WORD#16#8001 invalid measuringMode (PUB006); WORD#16#8002 hiLIM<=loLIM (PUB007).
Priority/simultaneous checks: measuringMode validity checked before hiLIM<=loLIM; simultaneous invalid mode and bad limits yields 16#8001 (unspecified, chosen).
outputValue: written only for enabled successful conversions; mode0 linear scaling clamped to 0/27648 or -27648/27648 (PUB003); mode1 raw/10 (PUB004); mode2 raw/100 (PUB005).
Read-only: analogValues unchanged; configuration fields only read (PUB001, PUB002).
Bounds: match by ordinal from each array lower bound; invalid count processes none.
Units: raw INT, output REAL, limits REAL; no time.
*)

(* CONTRACT_RULES [] *)

FUNCTION_BLOCK AnalogBatchProcessing
VAR_INPUT
    count : DINT;
END_VAR
VAR_IN_OUT
    analogValues : ARRAY[*] OF INT;
    channels : ARRAY[*] OF ST_AnalogChannel;
END_VAR
VAR
    tmp_lbA : DINT;
    tmp_lbC : DINT;
    tmp_availA : DINT;
    tmp_availC : DINT;
    tmp_process : DINT;
    tmp_i : DINT;
    tmp_idxA : DINT;
    tmp_idxC : DINT;
    tmp_raw : INT;
    tmp_rawReal : REAL;
    tmp_frac : REAL;
END_VAR

tmp_lbA := LOWER_BOUND(analogValues, 1);
tmp_lbC := LOWER_BOUND(channels, 1);
tmp_availA := UPPER_BOUND(analogValues, 1) - tmp_lbA + 1;
tmp_availC := UPPER_BOUND(channels, 1) - tmp_lbC + 1;

tmp_process := count;
IF tmp_process < 0 THEN
    tmp_process := 0;
END_IF;
IF tmp_process > tmp_availA THEN
    tmp_process := tmp_availA;
END_IF;
IF tmp_process > tmp_availC THEN
    tmp_process := tmp_availC;
END_IF;

FOR tmp_i := 0 TO tmp_process - 1 DO
    tmp_idxA := tmp_lbA + tmp_i;
    tmp_idxC := tmp_lbC + tmp_i;

    IF channels[tmp_idxC].enable THEN
        channels[tmp_idxC].retVal := WORD#0;

        IF (channels[tmp_idxC].measuringMode < 0) OR (channels[tmp_idxC].measuringMode > 2) THEN
            channels[tmp_idxC].retVal := WORD#16#8001;
            (* skip conversion; outputValue unchanged *)
        ELSIF channels[tmp_idxC].hiLIM <= channels[tmp_idxC].loLIM THEN
            channels[tmp_idxC].retVal := WORD#16#8002;
            (* skip conversion; outputValue unchanged *)
        ELSE
            tmp_raw := analogValues[tmp_idxA];
            tmp_rawReal := INT_TO_REAL(tmp_raw);

            CASE channels[tmp_idxC].measuringMode OF
                0:
                    IF channels[tmp_idxC].bipolar THEN
                        IF tmp_rawReal < -27648.0 THEN
                            tmp_rawReal := -27648.0;
                        ELSIF tmp_rawReal > 27648.0 THEN
                            tmp_rawReal := 27648.0;
                        END_IF;
                        tmp_frac := (tmp_rawReal + 27648.0) / 55296.0;
                    ELSE
                        IF tmp_rawReal < 0.0 THEN
                            tmp_rawReal := 0.0;
                        ELSIF tmp_rawReal > 27648.0 THEN
                            tmp_rawReal := 27648.0;
                        END_IF;
                        tmp_frac := tmp_rawReal / 27648.0;
                    END_IF;

                    channels[tmp_idxC].outputValue := channels[tmp_idxC].loLIM
                        + tmp_frac * (channels[tmp_idxC].hiLIM - channels[tmp_idxC].loLIM);

                1:
                    channels[tmp_idxC].outputValue := tmp_rawReal / 10.0;

                2:
                    channels[tmp_idxC].outputValue := tmp_rawReal / 100.0;

                ELSE
                    (* unreachable due to mode check above *)
                END_CASE;
        END_IF;
    END_IF;
END_FOR;

END_FUNCTION_BLOCK

(* ---- public-medium-02.candidate_02.st ---- *)
TYPE ST_AnalogChannel :
STRUCT
    enable : BOOL;
    hiLIM : REAL;
    loLIM : REAL;
    bipolar : BOOL;
    measuringMode : INT;
    retVal : WORD;
    outputValue : REAL;
END_STRUCT
END_TYPE;

(*
ENGINEERING_CONTRACT
Activation: process first count ordinal channels, count >= 0, clamped to min array lengths.
Enable: only channels[].enable = TRUE is evaluated; disabled rows retain previous retVal/outputValue.
retVal: for enabled rows write WORD#0 on success; WORD#16#8001 invalid measuringMode (PUB006); WORD#16#8002 hiLIM<=loLIM (PUB007).
Priority/simultaneous checks: measuringMode validity checked before hiLIM<=loLIM; simultaneous invalid mode and bad limits yields 16#8001 (unspecified, chosen).
outputValue: written only for enabled successful conversions; mode0 linear scaling clamped to 0/27648 or -27648/27648 (PUB003); mode1 raw/10 (PUB004); mode2 raw/100 (PUB005).
Read-only: analogValues unchanged; configuration fields only read (PUB001, PUB002).
Bounds: match by ordinal from each array lower bound; invalid count processes none.
Units: raw INT, output REAL, limits REAL; no time.
*)

(* CONTRACT_RULES [] *)

FUNCTION_BLOCK AnalogBatchProcessing
VAR_INPUT
    count : DINT;
END_VAR
VAR_IN_OUT
    analogValues : ARRAY[*] OF INT;
    channels : ARRAY[*] OF ST_AnalogChannel;
END_VAR
VAR
    tmp_lbA : DINT;
    tmp_lbC : DINT;
    tmp_availA : DINT;
    tmp_availC : DINT;
    tmp_process : DINT;
    tmp_i : DINT;
    tmp_idxA : DINT;
    tmp_idxC : DINT;
    tmp_raw : INT;
    tmp_rawReal : REAL;
    tmp_frac : REAL;
END_VAR

tmp_lbA := LOWER_BOUND(analogValues, 1);
tmp_lbC := LOWER_BOUND(channels, 1);
tmp_availA := UPPER_BOUND(analogValues, 1) - tmp_lbA + 1;
tmp_availC := UPPER_BOUND(channels, 1) - tmp_lbC + 1;

tmp_process := count;
IF tmp_process < 0 THEN
    tmp_process := 0;
END_IF;
IF tmp_process > tmp_availA THEN
    tmp_process := tmp_availA;
END_IF;
IF tmp_process > tmp_availC THEN
    tmp_process := tmp_availC;
END_IF;

FOR tmp_i := 0 TO tmp_process - 1 DO
    tmp_idxA := tmp_lbA + tmp_i;
    tmp_idxC := tmp_lbC + tmp_i;

    IF channels[tmp_idxC].enable THEN
        channels[tmp_idxC].retVal := WORD#0;

        IF (channels[tmp_idxC].measuringMode < 0) OR (channels[tmp_idxC].measuringMode > 2) THEN
            channels[tmp_idxC].retVal := WORD#16#8001;
            (* skip conversion; outputValue unchanged *)
        ELSIF channels[tmp_idxC].hiLIM <= channels[tmp_idxC].loLIM THEN
            channels[tmp_idxC].retVal := WORD#16#8002;
            (* skip conversion; outputValue unchanged *)
        ELSE
            tmp_raw := analogValues[tmp_idxA];
            tmp_rawReal := INT_TO_REAL(tmp_raw);

            CASE channels[tmp_idxC].measuringMode OF
                0:
                    IF channels[tmp_idxC].bipolar THEN
                        IF tmp_rawReal < -27648.0 THEN
                            tmp_rawReal := -27648.0;
                        ELSIF tmp_rawReal > 27648.0 THEN
                            tmp_rawReal := 27648.0;
                        END_IF;
                        tmp_frac := (tmp_rawReal + 27648.0) / 55296.0;
                    ELSE
                        IF tmp_rawReal < 0.0 THEN
                            tmp_rawReal := 0.0;
                        ELSIF tmp_rawReal > 27648.0 THEN
                            tmp_rawReal := 27648.0;
                        END_IF;
                        tmp_frac := tmp_rawReal / 27648.0;
                    END_IF;

                    channels[tmp_idxC].outputValue := channels[tmp_idxC].loLIM
                        + tmp_frac * (channels[tmp_idxC].hiLIM - channels[tmp_idxC].loLIM);

                1:
                    channels[tmp_idxC].outputValue := tmp_rawReal / 10.0;

                2:
                    channels[tmp_idxC].outputValue := tmp_rawReal / 100.0;

                ELSE
                    (* unreachable due to mode check above *)
                    tmp_raw := tmp_raw;   (* dummy statement to satisfy CASE syntax *)
                END_CASE;
        END_IF;
    END_IF;
END_FOR;

END_FUNCTION_BLOCK
